(* IEC 61131-3 sources: daoli-st-library/DL_Algo (part 21) *)

(* ---- FB_DL_SelfDischargeScreen.st ---- *)
(*
  FB_DL_SelfDischargeScreen  —  自放电筛分（压降速率 K 值分级 + 温度补偿） / Self-discharge screening by voltage-drop rate grading with temperature compensation
  分类 Category : DL_Algo
  版本 Version  : 1.0.0
  来源 Source   : roadmap-li-p2 — 锂电自放电筛分工站真缺口
  溯源 Origin   : 道莅 clean-room 实现；K 值 = ΔOCV/Δt 与 25 °C 温度补偿为公开自放电筛分算法，未复制任何源码行
  功能 Function : 1) 纯计算子函数 FC_DL_SelfDischargeKCalc 求压降速率
                  K = (fOcvStartV - fOcvEndV) / 静置时长(h)，静置时长按秒换算（除 3600.0 常量）；
                  2) 温度补偿：K25 = K / (1.0 + fTempCoeffPerK × (fTempC - 25.0))，
                  分母绝对值 <= 1.0E-6 返回 -1.0 哨兵（不饱和、不置 0，交主块判故障）；
                  3) 分级：K25 与 fClassAMvPerH / fClassBMvPerH / fClassCMvPerH 比较，
                  越 C 档为 eReject（ELSE 兜底）；
                  4) 报告值向上取整到 0.001 mV/h（先实数上限兜底 → 截断 → 余量进位，
                  正好整除不 +1，禁 TRUNC(x)+1）；
                  5) 本件只有故障码、无信息码（派单硬约束）。
  接口 Interface: 输入首末 OCV/静置时长/温度/温度系数/三档阈值；输出 K/K25/取整值/分级/码
  边界 Boundary : ① 组态闸：tRest <= T#0S、fTempCoeffPerK < 0.0、fClassAMvPerH < 0.0、
                  fClassBMvPerH <= fClassAMvPerH、fClassCMvPerH <= fClassBMvPerH
                  → 0389 锁存；② 首末 OCV 非有限（NaN 自反 + Inf 差值自减）→ 0389 锁存；
                  ③ 温补分母哨兵 -1.0 由主块转 0389 锁存（子函数不置故障）；
                  ④ 取整前实数上限兜底防 LREAL→DINT 溢出；⑤ 仅一个 R_TRIG，段 0 无条件调用；
                  ⑥ 故障相迁出唯一路径 = bReset 上升沿；⑦ 零全局耦合（无 GVL / %I %Q %M）。
  依赖 Depends  : Standard.library（R_TRIG）
  码表 Error codes（Algo 段 0002，故障窗口 0389；本件无信息码）:
    16#0002_0389 故障级：自放电筛分故障总码（组态非法 / OCV 非有限 / 温补分母非法），
                 锁存至 bReset 上升沿；归因见 eCause，不新增码位（派单硬约束单码）
  修订历史 Revision :
    2026-11-19  v1.0.0  R43 首版（批次 3 · 序号 13）
*)

TYPE E_DL_SdsState :
(
    eIdle   := 0,     // 未使能待筛分 / Idle, waiting screening
    eRun    := 10,    // 筛分计算中 / Screening active
    eFault  := 90     // 故障锁存相 / Fault latched phase
);
END_TYPE

TYPE E_DL_SdsClass :
(
    eNone   := 0,     // 未分级 / Not graded
    eClassA := 1,     // A 级（自放电最小） / Class A, lowest self-discharge
    eClassB := 2,     // B 级 / Class B
    eClassC := 3,     // C 级 / Class C
    eReject := 4      // 不合格（越 C 档） / Rejected
);
END_TYPE

TYPE E_DL_SdsCause :
(
    eNone       := 0, // 无故障成因 / No cause
    eCfgIllegal := 1, // 组态非法 / Illegal configuration
    eNonFinite  := 2, // OCV 非有限 / Non-finite OCV
    eCompDiv    := 3  // 温补分母非法 / Invalid compensation denominator
);
END_TYPE

FUNCTION FC_DL_SelfDischargeKCalc : REAL
VAR_INPUT
    fOcvStartV     : REAL;   // 静置前 OCV [V] / OCV before rest
    fOcvEndV       : REAL;   // 静置后 OCV [V] / OCV after rest
    fRestS         : REAL;   // 静置时长 [s]，域 > 0 / Rest duration in seconds
    fTempC         : REAL;   // 电芯温度 [°C] / Cell temperature
    fTempCoeffPerK : REAL;   // 温度系数 [1/K]，域 >= 0 / Temperature coefficient
END_VAR
VAR
    _fKPerH  : REAL;         // 未补偿压降速率 [V/h] / Uncompensated drop rate
    _fDen    : REAL;         // 温补分母 [-] / Compensation denominator
END_VAR
(* 纯计算子函数：K25 = K / (1 + coeff × (T - 25))；分母非法返回 -1.0 哨兵 *)
IF fRestS <= 1.0E-6 THEN                              // 除零前置判（时长正域） / Duration positive check
    FC_DL_SelfDischargeKCalc := -1.0;                 // 哨兵：时长非法 / Sentinel
    RETURN;
END_IF
_fKPerH := (fOcvStartV - fOcvEndV) / (fRestS / 3600.0);   // 压降速率 [V/h]（除常量 3600.0） / Drop rate
_fDen := 1.0 + fTempCoeffPerK * (fTempC - 25.0);          // 温补分母 / Compensation denominator
IF ABS(_fDen) <= 1.0E-6 THEN                          // 分母近零判据 / Near-zero denominator
    FC_DL_SelfDischargeKCalc := -1.0;                 // 哨兵：分母非法 / Sentinel
    RETURN;
END_IF
FC_DL_SelfDischargeKCalc := _fKPerH / _fDen * 1000.0; // 补偿后速率 [mV/h] / Compensated rate
END_FUNCTION

FUNCTION_BLOCK FB_DL_SelfDischargeScreen
VAR_INPUT
    fOcvStartV      : REAL := 0.0;      // 静置前 OCV [V] / OCV before rest
    fOcvEndV        : REAL := 0.0;      // 静置后 OCV [V] / OCV after rest
    tRest           : TIME := T#24H;    // 静置时长 [ms]，域 > 0 / Rest duration
    fTempC          : REAL := 25.0;     // 电芯温度 [°C] / Cell temperature
    fTempCoeffPerK  : REAL := 0.002;    // 温度系数 [1/K]，域 >= 0 / Temperature coefficient
    fClassAMvPerH   : REAL := 0.50;     // A 级上限 [mV/h] / Class A limit
    fClassBMvPerH   : REAL := 1.00;     // B 级上限 [mV/h] / Class B limit
    fClassCMvPerH   : REAL := 2.00;     // C 级上限 [mV/h] / Class C limit
    bEnable         : BOOL := FALSE;    // 筛分使能（电平）[-] / Screening enable
    bReset          : BOOL := FALSE;    // 复位命令，上升沿清故障 [-] / Reset edge
END_VAR
VAR_OUTPUT
    eState          : E_DL_SdsState;    // 状态出口，段 6 单点映射 / State outlet
    eClass          : E_DL_SdsClass;    // 分级出口 / Grading outlet
    eCause          : E_DL_SdsCause;    // 故障成因出口（R190） / Fault cause outlet
    fKMvPerH        : REAL;             // 温补后压降速率 [mV/h] / Compensated drop rate
    fKCeilMvPerH    : REAL;             // 向上取整到 0.001 的速率 [mV/h] / Ceiled rate
    bError          : BOOL;             // 故障锁存标志 [-] / Fault latch flag
    nErrId          : UDINT;            // 故障码，0 = 无故障（本件无信息码） / Fault code only
END_VAR
VAR
    _eState         : E_DL_SdsState := E_DL_SdsState.eIdle;   // 内部相位（CASE 唯一写入目标） / Internal phase
    _eClass         : E_DL_SdsClass := E_DL_SdsClass.eNone;   // 分级槽（每拍重算） / Grading slot
    _eCause         : E_DL_SdsCause := E_DL_SdsCause.eNone;   // 故障成因锁存（锁存量） / Latched cause
    rtReset         : R_TRIG;           // 复位沿实例，每周期无条件调用 / Reset edge
    _fK             : REAL;             // 子函数返回速率 [mV/h]（当拍量） / Sub-function result
    _fScaled        : REAL;             // 取整中间量（×1000 后） / Scaling intermediate
    _iScaled        : DINT;             // 截断后整数（×1000） / Truncated integer
    _bNonFin        : BOOL;             // OCV 非有限当拍量 [-] / Non-finite OCV
    _bCfgBad        : BOOL;             // 组态非法当拍量 [-] / Config illegal
    _bFault         : BOOL;             // 故障锁存位（锁存量） / Latched fault bit
    _uFault         : UDINT;            // 故障码锁存（锁存量） / Latched fault code
END_VAR

(* —— 段 0：沿实例无条件周期刷新 + 当拍量判据 —— *)
_bNonFin := (fOcvStartV <> fOcvStartV) OR (fOcvEndV <> fOcvEndV) OR (fTempC <> fTempC)
         OR ((fOcvStartV - fOcvStartV) <> (fOcvStartV - fOcvStartV))
         OR ((fOcvEndV - fOcvEndV) <> (fOcvEndV - fOcvEndV))
         OR ((fTempC - fTempC) <> (fTempC - fTempC));                        // NaN 自反 + Inf 差值自减 / NaN and Inf
_bCfgBad := (tRest <= T#0S) OR (fTempCoeffPerK < 0.0) OR (fClassAMvPerH < 0.0)
            OR (fClassBMvPerH <= fClassAMvPerH) OR (fClassCMvPerH <= fClassBMvPerH);   // 组态非法当拍量 / Config illegal
rtReset(CLK := bReset);                                                      // 复位沿，每拍必调 / Reset edge

(* —— 段 1：单拍量预清零（锁存量不入清单；分级槽每拍重算） —— *)
eClass := E_DL_SdsClass.eNone;      // 分级出口缺省未分级 / Grading default
fKMvPerH := 0.0;                    // 速率出口缺省 0 / Rate default
fKCeilMvPerH := 0.0;                // 取整出口缺省 0 / Ceil default
nErrId := 16#0000_0000;             // 故障码缺省无故障 / Fault code default

(* —— 段 2：复位沿 + 组态域闸 —— *)
IF rtReset.Q THEN                              // rtReset.Q = 当拍量 / current scan
    _bFault := FALSE;                          // 清故障锁存位（锁存量） / Clear fault latch
    _uFault := 16#0000_0000;                   // 清故障锁存码（锁存量） / Clear fault code
    _eCause := E_DL_SdsCause.eNone;            // 清成因（锁存量） / Clear cause
    IF _eState = E_DL_SdsState.eFault THEN
        _eState := E_DL_SdsState.eIdle;        // 故障相迁出：回未使能 / Fault exit to idle
    END_IF
END_IF
IF _bNonFin THEN                               // 非有限锁存 / Non-finite latch
    _uFault := 16#0002_0389;                   // 故障级：筛分故障总码 / Algo fault code
    _eCause := E_DL_SdsCause.eNonFinite;       // 归因：非有限 / Cause: non-finite
    _bFault := TRUE;                           // 标志与码位配对（R45） / Flag paired with code
END_IF
IF _bCfgBad THEN                               // 组态域闸 / Config gate
    _uFault := 16#0002_0389;
    _eCause := E_DL_SdsCause.eCfgIllegal;      // 归因：组态非法 / Cause: illegal config
    _bFault := TRUE;
END_IF

(* —— 段 3：K 值计算 + 温补哨兵 + 取整 + 分级（仅运行相且无故障） —— *)
IF (NOT _bFault) AND (_eState = E_DL_SdsState.eRun) THEN
    _fK := FC_DL_SelfDischargeKCalc(fOcvStartV := fOcvStartV, fOcvEndV := fOcvEndV,
                                    fRestS := TIME_TO_REAL(tRest) / 1000.0,
                                    fTempC := fTempC, fTempCoeffPerK := fTempCoeffPerK);   // 子函数求解（除零由子函数守卫） / Sub-function call
    IF _fK < 0.0 THEN                                      // 哨兵：时分母或时长非法 / Sentinel from sub-function
        _uFault := 16#0002_0389;
        _eCause := E_DL_SdsCause.eCompDiv;                 // 归因：温补分母非法 / Cause: denominator
        _bFault := TRUE;
    ELSE
        fKMvPerH := _fK;                                   // 速率镜像 / Rate mirror
        _fScaled := _fK * 1000.0;                           // 放大 1000 倍进入整数域 / Scale by thousand
        IF _fScaled >= 2.147483E9 THEN                      // 实数上限兜底（DINT 可表上界） / Real upper guard
            _fScaled := 2.147483E9;
        ELSIF _fScaled <= -2.147483E9 THEN                  // 实数下限兜底 / Real lower guard
            _fScaled := -2.147483E9;
        END_IF
        _iScaled := LREAL_TO_DINT(LREAL(_fScaled));         // 截断取整 / Truncate
        IF LREAL(_iScaled) < LREAL(_fScaled) - 1.0E-9 THEN  // 余量进位（正好整除不进位） / Ceiling by remainder
            _iScaled := _iScaled + 1;
        END_IF
        fKCeilMvPerH := DINT_TO_REAL(_iScaled) * 0.001;     // 还原为 0.001 mV/h 步长 / Restore 0.001 step
        IF fKCeilMvPerH <= fClassAMvPerH THEN
            _eClass := E_DL_SdsClass.eClassA;               // A 级 / Class A
        ELSIF fKCeilMvPerH <= fClassBMvPerH THEN
            _eClass := E_DL_SdsClass.eClassB;               // B 级 / Class B
        ELSIF fKCeilMvPerH <= fClassCMvPerH THEN
            _eClass := E_DL_SdsClass.eClassC;               // C 级 / Class C
        ELSE
            _eClass := E_DL_SdsClass.eReject;               // 不合格（ELSE 兜底） / Rejected fallback
        END_IF
    END_IF
END_IF

(* —— 段 4：故障解除式（R240；全当拍量）：rtReset.Q / NOT _bCfgBad / NOT _bNonFin —— *)
IF rtReset.Q AND (NOT _bCfgBad) AND (NOT _bNonFin) THEN
    _bFault := FALSE;                          // 清故障锁存位（锁存量） / Clear fault latch
    _uFault := 16#0000_0000;                   // 清故障锁存码（锁存量） / Clear fault code
    _eCause := E_DL_SdsCause.eNone;            // 清成因（锁存量） / Clear cause
END_IF

(* —— 段 4A：故障锁存相位迁移闸 —— *)
IF _bFault AND (_eState <> E_DL_SdsState.eFault) THEN
    _eState := E_DL_SdsState.eFault;           // 锁存即入故障相 / Latch enters fault phase
END_IF

(* —— 段 5：相位机（CASE 全覆盖 + ELSE 兜底） —— *)
CASE _eState OF

E_DL_SdsState.eIdle:
    IF bEnable AND (NOT _bFault) THEN          // 使能条件 / Enable gate
        _eState := E_DL_SdsState.eRun;         // 进筛分相 / Enter screening
    END_IF

E_DL_SdsState.eRun:
    IF NOT bEnable THEN                        // 撤使能：回未使能（前置消失） / Disable returns idle
        _eState := E_DL_SdsState.eIdle;
    END_IF

E_DL_SdsState.eFault:
    ;                                          // 故障相：仅段 4 复位沿可迁出 / Only reset exits

ELSE
    _uFault := 16#0002_0389;                   // 故障级：非法相位兜底（归并总码） / Illegal phase fallback
    _eCause := E_DL_SdsCause.eCfgIllegal;      // 归因：相位非法归并组态 / Cause: phase illegal
    _bFault := TRUE;
    _eState := E_DL_SdsState.eFault;           // 强制回故障相 / Force fault phase

END_CASE

(* —— 段 6：出口单点映射（名实同源；锁存码回放） —— *)
IF _bFault THEN
    nErrId := _uFault;                         // 故障锁存码回放 / Replay latched code
    eClass := E_DL_SdsClass.eNone;             // 故障相分级强制未分级 / Grading forced none
    fKCeilMvPerH := 0.0;                       // 故障相取整值强制 0（安全侧） / Ceil forced zero
ELSE
    nErrId := 16#0000_0000;                    // 无故障：本件无信息码 / No fault, no info code
    eClass := _eClass;                         // 分级出口 / Grading outlet
END_IF
bError := _bFault;                             // 故障标志同源 / Flag from latch
eState := _eState;                             // 状态出口 / State outlet
eCause := _eCause;                             // 成因出口 / Cause outlet

END_FUNCTION_BLOCK

(* ---- FB_DL_SensorConsensusSelector.st ---- *)
(*
  FB_DL_SensorConsensusSelector —— 多通道传感器共识选择：中位基准+偏差带剔除+通道不足降级到单通道，ENUM 状态机
  分类：DL_Algo | 复杂度：3 | 轮次：R86
  开源溯源：道莅原创（clean-room 自研，纯 IEC 61131-3 通用算法），无外部代码引用
  许可证：MIT

  职责：对 5 路同类传感器做共识表决——有效通道数 ≥3 时取中位数作基准、剔除超出偏差带的通道后取平均（NORMAL）；
        有效数 =2 取均值、=1 直通（DEGRADED）；有效数 =0 保持上值并置 xLost（LOST）。
  输入契约：arrVal 通道值 [工程单位]；arrValid 通道有效位；fDevBand 偏差带半宽 [工程单位]（> 0）；
            fAbsMax 非有限闸与量程闸的绝对上限 [工程单位]。
  输出契约：fOut 共识值 [工程单位]；nValidOut 参与表决的有效通道数；xValid 本次输出可信；
            xDegraded / xLost 分级标志；eMode 表决模式枚举。
  边界：① 非有限双判（x <> x 判 NaN、ABS(x) > fAbsMax 判 Inf / 越界）逐通道执行；
        ② 除零防护：所有均值前判分母 > 0；③ 排序用插入法（FOR + WHILE 递减），无 FOR..DOWNTO；
        ④ CASE 含 ELSE 兜底把非法模式拦入 LOST；⑤ 零全局耦合、零物理地址、零库件依赖。
*)

(*-----------------------------------------------------------------------------
 * 枚举: E_DL_ConsMode（共识表决模式，归属本文件，全库唯一定义）
 *----------------------------------------------------------------------------*)
TYPE E_DL_ConsMode :
(
    eNormal   := 0,   // 正常共识（≥3 通道且带内 ≥3） [—] / Normal consensus with at least three in band channels
    eDegraded := 1,   // 降级（2 通道均值 / 1 通道直通 / 带内不足 3） [—] / Degraded consensus
    eLost     := 2    // 失效（零有效通道，保持上值） [—] / Lost, holds the previous value
);
END_TYPE

FUNCTION_BLOCK FB_DL_SensorConsensusSelector
VAR_INPUT
    xEnable  : BOOL  := TRUE;                             // 使能，FALSE 时按失效模式处理 [—] / Enable, false is treated as lost
    arrVal   : ARRAY[0..4] OF REAL;                       // 五路通道采样值 [工程单位] / Five channel samples
    arrValid : ARRAY[0..4] OF BOOL;                       // 五路通道有效位 [—] / Five channel validity flags
    fDevBand : REAL  := 1.0;                              // 偏差带半宽，必须 > 0 [工程单位] / Deviation band half width
    fAbsMax  : REAL  := 1.0E30;                           // 数值绝对上限（非有限 / 越界闸） [工程单位] / The absolute magnitude gate
END_VAR
VAR_OUTPUT
    fOut       : REAL;                                    // 共识输出值 [工程单位] / The consensus output value
    nValidOut  : INT;                                     // 参与表决的有效通道数 [个] / The number of channels taking part
    xValid     : BOOL;                                    // 本次输出可信 [—] / The output is trustworthy
    xDegraded  : BOOL;                                    // 降级标志 [—] / The degraded flag
    xLost      : BOOL;                                    // 失效标志 [—] / The lost flag
    eMode      : E_DL_ConsMode;                           // 表决模式枚举 [—] / The consensus mode enumeration
END_VAR
VAR
    afSort    : ARRAY[0..4] OF REAL;                      // 有效值排序缓冲（升序） [工程单位] / The ascending sort buffer
    nCnt      : INT;                                      // 有效通道数 [个] / The valid channel count
    nIn       : INT;                                      // 偏差带内通道数 [个] / The in band channel count
    k         : INT;                                      // 外层遍历索引 [下标] / The outer loop index
    j         : INT;                                      // 插入排序内层索引 [下标] / The insertion sort index
    fTmp      : REAL;                                     // 插入排序暂存量 [工程单位] / The insertion sort temporary
    fMed      : REAL;                                     // 中位数基准 [工程单位] / The median reference
    fSum      : REAL;                                     // 带内累加和 [工程单位] / The in band accumulation
    fMean     : REAL;                                     // 带内均值 [工程单位] / The in band mean
    fCand     : REAL;                                     // 候选输出值 [工程单位] / The candidate output value
    fDiff     : REAL;                                     // 单通道与中位数的偏差 [工程单位] / The deviation from the median
    fLastOut  : REAL;                                     // 上拍共识输出保持量 [工程单位] / The held previous output
    xHasLast  : BOOL;                                     // 是否已有可用上拍值 [—] / Whether a previous value exists
    eCand     : E_DL_ConsMode;                            // 候选表决模式 [—] / The candidate mode
END_VAR
VAR CONSTANT
    DL_CM_ZERO : INT := 0;                                // 整型零常量 [个] / The integer zero constant
    DL_CM_ONE  : INT := 1;                                // 整型一常量 [个] / The integer one constant
    DL_CM_NCH  : INT := 5;                                // 通道总数 [个] / The total channel count
    DL_CM_MINC : INT := 3;                                // 正常共识所需最少通道数 [个] / The minimum channels for normal consensus
    DL_CM_R0   : REAL := 0.0;                             // 浮点零常量 [工程单位] / The floating point zero constant
    DL_CM_EPS  : REAL := 1.0E-6;                          // 浮点比较容差 [工程单位] / The floating point comparison tolerance
END_VAR

// 段 1｜输出预置（单点预置，CASE 之后不再无条件清零）
xValid := FALSE;                                          // 可信位预置假 / preset the valid flag false
xDegraded := FALSE;                                       // 降级位预置假 / preset the degraded flag false
xLost := FALSE;                                           // 失效位预置假 / preset the lost flag false
nValidOut := DL_CM_ZERO;                                  // 有效通道数预置零 [个] / preset the valid count zero
nCnt := DL_CM_ZERO;                                       // 排序缓冲计数预置零 [个] / preset the buffer count zero
fMed := DL_CM_R0;                                         // 中位数预置零 [工程单位] / preset the median zero
fCand := fLastOut;                                        // 候选值默认继承上拍值 [工程单位] / default the candidate to the held value

// 段 2｜逐通道有效性 + 非有限闸，有效值收集进排序缓冲
FOR k := DL_CM_ZERO TO DL_CM_NCH - 1 DO                   // 五通道遍历（上界 4 已由常量钉死） / traverse all channels
    IF arrValid[k] THEN                                   // 通道有效位为真 / the channel is flagged valid
        IF (arrVal[k] <> arrVal[k]) THEN                  // 自反判 NaN / the self comparison catches NaN
            fTmp := DL_CM_R0;                             // 置暂存零（本通道将被剔除） / stage zero, channel dropped
        ELSIF ABS(arrVal[k]) > fAbsMax THEN               // 越绝对上限判 Inf / 越界 / beyond the magnitude gate
            fTmp := DL_CM_R0;                             // 置暂存零（本通道将被剔除） / stage zero, channel dropped
        ELSE
            afSort[nCnt] := arrVal[k];                    // 有效值入缓冲 [工程单位] / store the valid value
            nCnt := nCnt + DL_CM_ONE;                     // 有效计数自增 [个] / increment the valid count
        END_IF
    END_IF
END_FOR
nValidOut := nCnt;                                        // 有效通道数出口 [个] / publish the valid count

// 段 3｜插入排序升序（WHILE 显式递减，禁 FOR..DOWNTO）
FOR k := DL_CM_ONE TO nCnt - DL_CM_ONE DO                 // 从第二个元素起逐个插入 / insert every element from the second
    IF k >= DL_CM_ONE THEN                                // k 合法且缓冲至少有 k+1 个元素 / k is legal with enough elements
        fTmp := afSort[k];                                // 取出待插入元素 [工程单位] / take the element to insert
        j := k - DL_CM_ONE;                               // 内层索引从 k-1 起 / the inner index starts at k minus one
        WHILE (j >= DL_CM_ZERO) AND (afSort[j] > fTmp) DO // 显式递减并判下界 / explicit decrement with a bound check
            afSort[j + DL_CM_ONE] := afSort[j];           // 逆序元素右移一格 / shift the larger element right
            j := j - DL_CM_ONE;                           // 内层索引递减 [下标] / decrement the inner index
        END_WHILE
        afSort[j + DL_CM_ONE] := fTmp;                    // 待插入元素落位 [工程单位] / land the element
    END_IF
END_FOR

// 段 4｜按有效通道数分档：中位数基准 + 偏差带剔除 + 候选模式判定
IF (NOT xEnable) OR (nCnt = DL_CM_ZERO) THEN              // 未使能或零有效通道 / disabled or no valid channel
    eCand := E_DL_ConsMode.eLost;                         // 候选模式判失效 / the candidate mode is lost
ELSIF nCnt = DL_CM_ONE THEN                               // 单通道直通 / a single channel passes through
    fCand := afSort[0];                                   // 直通该通道值 [工程单位] / pass the single value
    eCand := E_DL_ConsMode.eDegraded;                     // 候选模式判降级 / the candidate mode is degraded
ELSIF nCnt = DL_CM_ONE + DL_CM_ONE THEN                   // 双通道取均值 / two channels take the mean
    fCand := (afSort[0] + afSort[1]) / 2.0;               // 双通道均值 [工程单位] / the mean of the two channels
    eCand := E_DL_ConsMode.eDegraded;                     // 候选模式判降级 / the candidate mode is degraded
ELSE                                                      // 三通道及以上做中位基准表决 / three or more channels vote
    IF (nCnt MOD 2) = DL_CM_ONE THEN                      // 奇数个取正中位 / odd count takes the middle element
        fMed := afSort[nCnt / 2];                         // 中位数基准 [工程单位] / the median reference
    ELSE
        fMed := (afSort[nCnt / 2 - DL_CM_ONE] + afSort[nCnt / 2]) / 2.0; // 偶数个取中间两值均值 [工程单位]
    END_IF
    nIn := DL_CM_ZERO;                                    // 带内计数清零 [个] / clear the in band count
    fSum := DL_CM_R0;                                     // 带内和清零 [工程单位] / clear the in band sum
    FOR k := DL_CM_ZERO TO nCnt - DL_CM_ONE DO             // 遍历有效通道做偏差带剔除 / filter by the deviation band
        fDiff := afSort[k] - fMed;                        // 与中位数的偏差 [工程单位] / the deviation from the median
        IF ABS(fDiff) <= fDevBand THEN                    // 带内（含边界，容差口径） / inside the band
            fSum := fSum + afSort[k];                     // 累加带内值 [工程单位] / accumulate the in band value
            nIn := nIn + DL_CM_ONE;                       // 带内计数自增 [个] / increment the in band count
        END_IF
    END_FOR
    IF nIn >= DL_CM_MINC THEN                             // 带内至少 3 通道 / at least three channels stay in band
        fMean := fSum / INT_TO_REAL(nIn);                 // 带内均值（分母 ≥3 已证非零） [工程单位] / the in band mean
        fCand := fMean;                                   // 候选输出取带内均值 [工程单位] / the candidate is the mean
        eCand := E_DL_ConsMode.eNormal;                    // 候选模式判正常 / the candidate mode is normal
    ELSIF nIn = DL_CM_ONE + DL_CM_ONE THEN                // 带内仅剩 2 通道 / only two channels stay in band
        fMean := fSum / 2.0;                              // 两通道均值 [工程单位] / the mean of the two channels
        fCand := fMean;                                   // 候选输出取该均值 [工程单位] / the candidate is that mean
        eCand := E_DL_ConsMode.eDegraded;                 // 候选模式判降级 / the candidate mode is degraded
    ELSE                                                  // 带内不足 2 通道，退回中位基准 / too few in band, fall back to the median
        fCand := fMed;                                    // 候选输出取中位数 [工程单位] / the candidate is the median
        eCand := E_DL_ConsMode.eDegraded;                 // 候选模式判降级 / the candidate mode is degraded
    END_IF
END_IF

// 段 5｜模式出口分派（ENUM + CASE，ELSE 拦截非法模式）
CASE eCand OF
    E_DL_ConsMode.eNormal:
        fOut := fCand;                                    // 正常模式直接输出候选值 [工程单位] / publish the candidate
        xValid := TRUE;                                   // 置可信位 [—] / raise the valid flag
        xDegraded := FALSE;                               // 清降级位 [—] / clear the degraded flag
        xLost := FALSE;                                   // 清失效位 [—] / clear the lost flag
        fLastOut := fOut;                                 // 刷新保持量 [工程单位] / refresh the held value
        xHasLast := TRUE;                                 // 保持量可用 [—] / the held value is now available
    E_DL_ConsMode.eDegraded:
        fOut := fCand;                                    // 降级模式输出候选值 [工程单位] / publish the candidate
        xValid := TRUE;                                   // 降级输出仍可信 [—] / a degraded output is still valid
        xDegraded := TRUE;                                // 置降级位 [—] / raise the degraded flag
        xLost := FALSE;                                   // 清失效位 [—] / clear the lost flag
        fLastOut := fOut;                                 // 刷新保持量 [工程单位] / refresh the held value
        xHasLast := TRUE;                                 // 保持量可用 [—] / the held value is now available
    E_DL_ConsMode.eLost:
        IF xHasLast THEN                                  // 已有上拍值 / a previous value exists
            fOut := fLastOut;                             // 保持上拍值 [工程单位] / hold the previous value
        ELSE
            fOut := DL_CM_R0;                             // 无上拍值输出零哨兵 [工程单位] / zero sentinel without history
        END_IF
        xValid := FALSE;                                  // 失效输出不可信 [—] / the lost output is not valid
        xDegraded := TRUE;                                // 失效同时视为降级 [—] / lost is also degraded
        xLost := TRUE;                                    // 置失效位 [—] / raise the lost flag
ELSE
    fOut := DL_CM_R0;                                     // 非法模式输出零哨兵 [工程单位] / illegal mode outputs the zero sentinel
    xValid := FALSE;                                      // 非法模式不可信 [—] / an illegal mode is not valid
    xDegraded := TRUE;                                    // 非法模式视为降级 [—] / an illegal mode is degraded
    xLost := TRUE;                                        // 非法模式视为失效 [—] / an illegal mode is lost
    eCand := E_DL_ConsMode.eLost;                          // 非法模式回写为失效 [—] / normalise the illegal mode to lost
END_CASE
eMode := eCand;                                           // 模式枚举单点出口 / the single point mode outlet
END_FUNCTION_BLOCK

(* ---- FB_DL_SensorDriftBaseline.st ---- *)
(*
  Name        : FB_DL_SensorDriftBaseline
  Category    : DL_Algo
  Version     : 1.0.1
  Purpose     : 传感器慢漂移基线跟踪：长窗指数（EMA）基线随测量缓慢跟随，测量对基线的快偏差超限经确认延时即报警（区分真实工况阶跃与传感器漂移）；/ Sensor slow-drift baseline tracking: a long-window EMA baseline follows the measurement, and a fast deviation beyond limit confirmed over a delay raises an alarm
  溯源        : 借 t2-1-measurement 的分类/参数域组织，clean-room 实现
  Changelog   : v1.0.1 R54 非有限输入穿透修复：迁入拍/基线更新/残差出口前置有限性闸，非有限拍冻结基线并置 bSensorBad，出口保持上拍值
  Boundary    : ① 组态闸：基线因子域 (0..1] / 快偏差限 > 0 / 确认延时 > 0 → 锁存故障（因子 0/1 端点使基线冻结或退化为直通）；
                ② 非有限测量该拍不更新基线（基线保持上拍值，防污染慢积分器），判据整拍跳过；
                ③ 基线快照在迁入 eMon 拍取（fValue 首值），避免从 0 慢爬造成的假偏差；
                ④ 确认延时 TON 串 eMon 相位闸（族③），段 0 无 IF 包裹；
                ⑤ bDriftFast 锁存至复位沿；fBaseline/fDeviation 出口在 eIdle/eFault 有确定值；
                ⑥ 本件为诊断层，不修正测量值、不重标定（属主边界）。
*)
TYPE E_DL_SdbState :
(
    eIdle  := 0,                             (* 未使能 / Disabled *)
    eMon   := 10,                            (* 基线跟踪运行 / Tracking *)
    eFault := 90                             (* 故障锁存相 / Fault latched *)
);
END_TYPE

TYPE E_DL_SdbCause :
(
    eNone       := 0,                        (* 无故障成因 / No cause *)
    eCfgIllegal := 1,                        (* 组态非法：因子/偏差限/延时越域 / Illegal config *)
    eDriftFast  := 2,                        (* 快偏差确认（基线失跟或真实阶跃，上层判别） / Fast deviation confirmed *)
    ePhaseBad   := 3                         (* 非法相位兜底 / Illegal phase fallback *)
);
END_TYPE

FUNCTION_BLOCK FB_DL_SensorDriftBaseline
VAR_INPUT
    fValue    : REAL := 0.0;                 (* 传感器测量值（任意工程量）[-] / Sensor measurement *)
    fAlpha    : REAL := 0.005;               (* 基线 EMA 因子（每拍跟随比例），域 (0..1] [-] / Baseline EMA factor *)
    fFastLim  : REAL := 5.0;                 (* 快偏差报警限，域 > 0 [工程单位] / Fast-deviation limit, > 0 *)
    tConfirm  : TIME := T#30S;               (* 快偏差确认延时，域 > T#0S [ms] / Deviation confirm delay, > 0 *)
    bEnable   : BOOL := TRUE;                (* 跟踪使能 [-] / Enable *)
    bReset    : BOOL := FALSE;               (* 复位命令，上升沿清报警与基线 [-] / Reset command *)
END_VAR
VAR_OUTPUT
    fBaseline : REAL;                        (* 慢漂移基线（EMA 跟踪值）[工程单位] / Slow-drift baseline *)
    fDeviation: REAL;                        (* 测量对基线快偏差（实时派生）[工程单位] / Fast deviation versus baseline *)
    bDriftFast: BOOL;                        (* 快偏差报警锁存（复位沿清）[-] / Fast-deviation alarm latched *)
    bSensorBad: BOOL;                        (* 测量非有限传感器失效锁存（复位沿清，v1.0.1）[-] / Sensor bad latched *)
    eState    : E_DL_SdbState;               (* 状态出口 / State outlet *)
    eCause    : E_DL_SdbCause;               (* 故障成因出口（R190 归因唯一） / Fault cause outlet *)
    bError    : BOOL;                        (* 故障锁存标志 [-] / Fault latch flag *)
END_VAR
VAR
    _eState  : E_DL_SdbState := E_DL_SdbState.eIdle;     (* 内部相位（CASE 唯一写入目标） / Internal phase *)
    _eCause  : E_DL_SdbCause := E_DL_SdbCause.eNone;     (* 故障成因锁存量 / Latched cause *)
    rtReset  : R_TRIG;                       (* 复位沿实例，段 0 无条件调用 / Reset edge instance *)
    tonConf  : TON;                          (* 快偏差确认延时计时器（IN 由偏差判据派生 + 相位闸） / Deviation confirm timer *)
    _bFault  : BOOL;                         (* 故障锁存位 / Latched fault bit *)
    _bCfgBad : BOOL;                         (* 组态非法当拍量 / Illegal config this scan *)
    _bFin    : BOOL;                         (* 测量值有限性当拍量 / Measurement finiteness *)
    _bBase   : BOOL;                         (* 基线已建立标志 / Baseline established flag *)
    _fBaseI  : REAL;                         (* 基线内部量（EMA 状态）[工程单位] / Baseline internal EMA state *)
    _fDevI   : REAL;                         (* 快偏差中间量 [工程单位] / Deviation intermediate *)
    _fDevLast: REAL;                         (* 上拍有效偏差快照（非有限拍出口冻结用，v1.0.1）[工程单位] / Last valid deviation snapshot *)
    _bDevRaw : BOOL;                         (* 快偏差原始判据当拍量 / Raw deviation verdict *)
END_VAR
VAR CONSTANT
    DL_SDB_EPS  : REAL := 1.0E-6;            (* 判零容差 [-] / Epsilon *)
    DL_SDB_ONE  : REAL := 1.0;               (* 因子上界常量 [-] / Factor upper bound *)
END_VAR

(* —— 段 0：当拍判据派生 + 实例无条件刷新（R228A；R_TRIG/TON 全在段 0，无 IF 包裹） —— *)
_bCfgBad := (fAlpha <= DL_SDB_EPS) OR (fAlpha > DL_SDB_ONE)                    (* 基线因子域闸 (0..1]（端点退化解拦截） / Factor domain gate *)
            OR (fFastLim <= DL_SDB_EPS)                                        (* 快偏差限正域闸 / Deviation limit gate *)
            OR NOT (tConfirm > T#0S);                                          (* 确认延时正域闸 / Confirm delay gate *)
rtReset(CLK := bReset);                                                        (* 复位沿每拍必调 / Reset edge every scan *)
_bFin := (fValue = fValue) AND ((fValue - fValue) = (fValue - fValue));        (* 测量值 NaN 自反 + Inf 差判闸 / Measurement NaN and Inf gate *)
_fDevI := 0.0;                                                                 (* 偏差中间量预置（基线无效期为 0，不误触发计时） / Deviation preset zero *)
IF _bFin AND _bBase THEN
    _fDevI := fValue - _fBaseI;                                                (* 快偏差 = 测量 - 基线（基线已建立才派生）[工程单位] / Deviation versus baseline *)
END_IF
_bDevRaw := _bFin AND _bBase AND (ABS(_fDevI) > fFastLim);                     (* 原始判据：有限 + 基线在 + 超限（直比阈值，非浮点等值） / Raw deviation verdict *)
tonConf(IN := (_eState = E_DL_SdbState.eMon) AND _bDevRaw, PT := tConfirm);    (* 确认延时：判据持续才计时，串 eMon 相位闸 / Confirm timer with phase gate *)

(* —— 段 1：单拍量预清零（R107；bDriftFast 为锁存出口不预清，复位沿清，族② 口径） —— *)
fBaseline := 0.0;                                                              (* 基线出口预清（派生拍覆盖） / Baseline outlet preset *)
fDeviation := 0.0;                                                             (* 偏差出口预清 / Deviation outlet preset *)

(* —— 段 2：复位沿处理（作用域：清故障 + 清报警 + 清基线 + 迁 eIdle，R283 逐项声明） —— *)
IF rtReset.Q THEN
    _bFault := FALSE;                                                          (* 清故障锁存 / Clear fault *)
    _eCause := E_DL_SdbCause.eNone;                                            (* 清成因 / Clear cause *)
    bDriftFast := FALSE;                                                       (* 清快偏差报警锁存 / Clear alarm latch *)
    _bBase := FALSE;                                                           (* 清基线已建立位（重使能重新取快照） / Clear baseline flag *)
    _fBaseI := 0.0;                                                            (* 清基线内部量 / Clear baseline internal *)
    _fDevLast := 0.0;                                                          (* 清有效偏差快照（v1.0.1） / Clear deviation snapshot *)
    bSensorBad := FALSE;                                                       (* 清传感器失效锁存（v1.0.1） / Clear sensor bad latch *)
    fBaseline := 0.0;                                                          (* 清基线出口 / Clear baseline outlet *)
    fDeviation := 0.0;                                                         (* 清偏差出口 / Clear deviation outlet *)
    _eState := E_DL_SdbState.eIdle;                                            (* 迁未使能相 / Back to idle *)
END_IF

(* —— 段 3：组态故障锁存（锁存至复位沿，R189） —— *)
IF _bCfgBad AND NOT _bFault THEN
    _bFault := TRUE;                                                           (* 锁存故障位 / Latch fault *)
    _eCause := E_DL_SdbCause.eCfgIllegal;                                      (* 成因：组态非法 / Cause: illegal config *)
    _eState := E_DL_SdbState.eFault;                                           (* 同步迁故障相 / Migrate to fault *)
END_IF

(* —— 段 4：CASE 主状态机（ELSE 兜底迁 eFault，红线 6） —— *)
CASE _eState OF
    E_DL_SdbState.eIdle:                                                       (* 未使能：出口确定值 / Disabled *)
        fBaseline := 0.0;                                                      (* 失能清基线出口 / Clear baseline outlet *)
        fDeviation := 0.0;                                                     (* 失能清偏差出口 / Clear deviation outlet *)
        bDriftFast := FALSE;                                                   (* 失能清报警出口 / Clear alarm outlet *)
        _bBase := FALSE;                                                       (* 失能清基线位（重使能重新对齐） / Clear baseline flag *)
        bSensorBad := FALSE;                                                   (* 失能清传感器失效出口（确定值） / Clear sensor bad *)
        IF bEnable AND NOT _bFault AND _bFin THEN                              (* 迁入闸加有限性闸：迁入拍为非有限不建基线不迁入（v1.0.1 修复） / Entry gate with finiteness *)
            _fBaseI := fValue;                                                 (* 迁入拍取基线首快照（相位闸配套，边界③） / Baseline snapshot at entry *)
            _bBase := TRUE;                                                    (* 基线已建立 / Baseline established *)
            _eState := E_DL_SdbState.eMon;                                     (* 使能进入跟踪 / Enter tracking *)
        END_IF
    E_DL_SdbState.eMon:                                                        (* 跟踪相：EMA 基线 + 快偏差判 / Tracking *)
        IF NOT bEnable THEN
            _eState := E_DL_SdbState.eIdle;                                    (* 失能回未使能 / Back to idle *)
        ELSE
            fBaseline := _fBaseI;                                              (* 基线出口（状态镜像，R191；非有限拍 _fBaseI 冻结即保持上拍） / Baseline outlet *)
            IF _bFin THEN
                fDeviation := _fDevI;                                          (* 偏差出口（有限拍派生） / Deviation outlet *)
                _fDevLast := _fDevI;                                           (* 有效偏差快照推进（v1.0.1） / Advance deviation snapshot *)
                _fBaseI := _fBaseI + fAlpha * (fValue - _fBaseI);              (* EMA 基线慢跟随（因子域闸保证 (0..1]） / EMA baseline update *)
            ELSE
                fDeviation := _fDevLast;                                       (* 非有限拍：偏差出口保持上拍值（v1.0.1 修复） / Hold last deviation *)
                bSensorBad := TRUE;                                            (* 非有限拍置传感器失效锁存（复位沿清，v1.0.1） / Sensor bad latch *)
            END_IF
            IF tonConf.Q THEN                                                  (* 快偏差持续满确认延时：报警 / Deviation confirmed *)
                bDriftFast := TRUE;                                            (* 报警锁存（复位沿清） / Latch alarm *)
                _bFault := TRUE;                                               (* 同步故障锁存（R45 配对） / Latch fault *)
                _eCause := E_DL_SdbCause.eDriftFast;                           (* 成因：快偏差 / Cause: fast deviation *)
            END_IF
        END_IF
    E_DL_SdbState.eFault:                                                      (* 故障相：冻结保持末值，仅复位沿出 / Fault *)
        ;                                                                      (* 锁存回放（R28） / Replay from latch *)
    ELSE                                                                       (* 非法相位兜底迁安全态 / Illegal phase fallback *)
        _eState := E_DL_SdbState.eFault;                                       (* 迁故障相 / To fault *)
        _bFault := TRUE;                                                       (* 同步锁存 / Latch *)
        _eCause := E_DL_SdbCause.ePhaseBad;                                    (* 成因：非法相位 / Cause: illegal phase *)
END_CASE

(* —— 段 5：出口映射（bError/eState 同源，R191） —— *)
bError := _bFault;                                                             (* 故障标志镜像 / Fault flag mirror *)
eState := _eState;                                                             (* 状态出口 / State outlet *)
eCause := _eCause;                                                             (* 成因出口 / Cause outlet *)
END_FUNCTION_BLOCK

(* ---- FB_DL_SensorFusion2.st ---- *)
(*==============================================================================
 * 组件名称 (Component)  : FB_DL_SensorFusion2
 * 所属子库 (Sublibrary) : DL_Algo
 * 当前版本 (Version)    : 1.0.1
 * 兼容性   (Platform)   : CODESYS 3.5+ / TwinCAT 3 / 汇川 InoProShop / 施耐德 Machine Expert
 *                         仅依赖 Standard.library（ABS），零厂商私有库
 * 功能描述 (Function)   : 双传感器方差加权融合：对同一物理量的两路测量（如 RTD+红外温漂
 *                         互补型双测）按在线递推噪声方差倒数动态配权：
 *                           _fVarX := (1-fTauVar)×_fVarX + fTauVar×(fMeasX-_fMean)²
 *                           fWeightA = (1/_fVarA) / ((1/_fVarA)+(1/_fVarB))
 *                           fFused   = fWeightA×fMeasA + (1-fWeightA)×fMeasB
 *                         一致性判据 bAgree = |fMeasA-fMeasB| <= fDevMax；单源失效全权重
 *                         交给健康源（降级不拒算）；双源失效冻结上次 fFused 且 bValid=FALSE。
 * 接口     (Interface)  : 输入 fMeasA/fMeasB 双路测量、bFreshA/bFreshB 数据新鲜度、
 *                         fTauVar 方差递推平滑系数（域 0~1 无量纲）、fDevMax 一致性偏差闸
 *                         （工程单位）、bReset 复位；输出 fFused 融合值、fWeightA 权重
 *                         （0~1）、bAgree 一致性、bValid 有效标志、bError 故障标志。
 * 边界     (Boundary)   : ① **属主边界（写死）：本件只做双源静态融合，不判传感器硬故障、
 *                         不切换通道、不接管信号健康诊断**；通道硬失效裁决归
 *                         `FB_DL_RedundantSwitch`（二选一切换），本件是"都信、按噪声配权"。
 *                         ② 方差下限钳 fVarMin（VAR CONSTANT）防除零：权重分母两项各含
 *                         1/_fVarX，钳底后分母恒正，无需额外除零判。
 *                         ③ 非有限值当拍剔除（R245）：该源当拍视同不新鲜；双源当拍均剔除
 *                         → 冻结 fFused、bValid=FALSE。
 *                         ④ 权重输出钳 [0,1]；fTauVar 组态域闸（<0 或 >1）与 fDevMax<0
 *                         → 锁存 bError，冻结输出，解除沿 = bReset 上升沿。
 *                         ⑤ 方差递推仅在双源同拍有效时进行（单源降级只直通，不污染方差）。
 *                         ⑥ 零全局耦合（无 GVL / 无 VAR_EXTERNAL / 无物理地址）。
 * 分工声明 (Scope)      : 与 `FB_DL_KalmanFilter1D` 分工：单流递推滤波 ≠ 双源加权融合；
 *                         与 `FB_DL_RedundantSwitch` 分工：二选一切换 ≠ 加权融合（见①）。
 * 来源标签 (Source Tag) : 自研线（公开加权融合公式 clean-room，逆方差权重为公开统计定义）
 * 码表     (Codes)      : 本件不占用任何全局数字码位。出口为 LREAL 组 + BOOL 组；
 *                         数字码位待主控收口阶段统一派号。
 * 红线自检 (Redline)    : R1 ✓ 零 GVL/VAR_EXTERNAL ｜ R2 ✓ 零 %I/%Q/%M ｜ R3 ✓ 纯 IEC 61131-3
 *                         R4 ✓ 方差下限防除零 + 非有限剔除 + 权重钳位 ｜ R5 ✓ 声明逐行同行双语注释
 *                         R6 N/A（无 ENUM 状态机） ｜ R7 ✓ 一 R_TRIG 段 0 无条件刷新
 * 修订历史 (Revision)   : 2026-11-20  v1.0.1  R50 返修 R3：fTauVar=0 端点防护
 *                         （下限钳位）——fTauVar=0 时方差递推步长为零，方差
 *                         永冻结于初值 1.0、权重恒 0.5（自适应失效），现引入
 *                         DL_SF2_TAUMIN(1E-6) 下限钳位使递推保持最低活跃度；
 *                         行为变更同步更新验收向量（fTauVar=0 按 1E-6 生效）。
 *                         2026-11-20  v1.0.0  R48 首版（批次 2 · 序号 6）
 *                         验收向量：等方差双源 → 权重 0.5；A 方差骤增 → 权重移向 B；
 *                         A 不新鲜 → 权重 1.0 全信 B；双源失效 → 冻结 + bValid=FALSE。
 *==============================================================================*)

FUNCTION_BLOCK FB_DL_SensorFusion2
VAR_INPUT
    fMeasA  : LREAL := 0.0;    // A 源测量值 [工程单位] / Source A measurement
    fMeasB  : LREAL := 0.0;    // B 源测量值（与 A 同物理量） [工程单位] / Source B measurement, same quantity as A
    bFreshA : BOOL := TRUE;    // A 源数据新鲜度 [-] / Source A freshness
    bFreshB : BOOL := TRUE;    // B 源数据新鲜度 [-] / Source B freshness
    fTauVar : LREAL := 0.1;    // 方差递推平滑系数，域 [0,1] [无量纲] / Variance recursion smoothing factor
    fDevMax : LREAL := 1.0;    // 一致性偏差闸（|A-B| 超此值 bAgree=FALSE） [工程单位] / Agreement deviation gate
    bReset  : BOOL := FALSE;   // 复位，上升沿清组态故障锁存 [-] / Reset, rising edge clears config fault
END_VAR
VAR_OUTPUT
    fFused   : LREAL;          // 融合输出值 [工程单位] / Fused output value
    fWeightA : LREAL;          // A 源权重，域 [0,1] [-] / Source A weight in [0,1]
    bAgree   : BOOL;           // 双源一致性（单源降级恒 TRUE） [-] / Two-source agreement
    bValid   : BOOL;           // 融合有效标志（双源失效/组态故障为 FALSE） [-] / Fusion validity flag
    bError   : BOOL;           // 组态故障标志（锁存） [-] / Configuration fault flag, latched
END_VAR
VAR
    _fVarA    : LREAL := 1.0;  // A 源在线递推噪声方差（初值 1.0，量纲平方） / Source A recursive noise variance
    _fVarB    : LREAL := 1.0;  // B 源在线递推噪声方差（初值 1.0） / Source B recursive noise variance
    _fMean    : LREAL := 0.0;  // 上拍融合均值（方差递推参考点，冻结源） / Previous fused mean, recursion reference
    _fW       : LREAL := 0.5;  // 当拍权重中间量（冻结源，与出口同源） / Weight intermediate, frozen source
    _fTauUse  : LREAL;         // 生效递推系数（下限钳位后，v1.0.1 端点防护） [-] / Effective smoothing factor after floor clamp
    _fFused   : LREAL := 0.0;  // 融合值锁存镜像（冻结语义源） / Fused value latch mirror
    _bValid   : BOOL;          // 有效标志内部量 / Validity internal
    _bErrLatch: BOOL;          // 组态故障锁存位（解除沿 = bReset 上升沿） / Latched config fault, cleared by reset edge
    rtReset   : R_TRIG;        // 复位沿实例，段 0 无条件调用 / Reset edge instance
    _bUseA    : BOOL;          // A 源当拍可用（新鲜 ∧ 有限） / Source A usable this scan
    _bUseB    : BOOL;          // B 源当拍可用 / Source B usable this scan
    _fInvA    : LREAL;         // A 源逆方差中间量 / Inverse variance of A
    _fInvB    : LREAL;         // B 源逆方差中间量 / Inverse variance of B
    _fDevA    : LREAL;         // A 源对均值偏差 [工程单位] / Deviation of A from mean
    _fDevB    : LREAL;         // B 源对均值偏差 [工程单位] / Deviation of B from mean
END_VAR
VAR CONSTANT
    DL_SF2_VARMIN : LREAL := 1.0E-12;   // 方差下限钳（防除零） [工程单位²] / Variance floor against zero division
    DL_SF2_TAUMIN : LREAL := 1.0E-6;    // 递推系数下限钳（fTauVar=0 端点防护，v1.0.1） [-] / Smoothing factor floor, endpoint guard
    DL_SF2_EPS    : LREAL := 0.0;       // 非有限差值判零基准 [-] / Non-finite difference zero base
    DL_SF2_ONE    : LREAL := 1.0;       // 单位常量（权重钳上限） [-] / Unit constant, weight ceiling
END_VAR

(* —— 段 0：非有限判 + 组态闸 + 沿刷新 —— *)
_bUseA := bFreshA AND (fMeasA = fMeasA) AND ((fMeasA - fMeasA) = DL_SF2_EPS);   // A 源新鲜 ∧ 有限（NaN 自不等 / Inf 差非零，R245） / A fresh and finite
_bUseB := bFreshB AND (fMeasB = fMeasB) AND ((fMeasB - fMeasB) = DL_SF2_EPS);   // B 源新鲜 ∧ 有限 / B fresh and finite
IF (fTauVar < 0.0) OR (fTauVar > DL_SF2_ONE) OR (fDevMax < 0.0) THEN
    _bErrLatch := TRUE;                                    // 组态域闸：锁存（R188 解除沿 = bReset 上升沿） / Config domain gate: latch
END_IF
_fTauUse := fTauVar;                                       // 生效递推系数工作副本 / Effective factor working copy
IF _fTauUse < DL_SF2_TAUMIN THEN
    _fTauUse := DL_SF2_TAUMIN;                             // fTauVar=0 端点钳位：递推保持最低活跃度（v1.0.1） / Endpoint floor clamp
END_IF
rtReset(CLK := bReset);                                    // 复位沿，每拍必调 / Reset edge, every scan

(* —— 段 1：复位沿 —— *)
IF rtReset.Q THEN
    _bErrLatch := FALSE;                                   // 清组态故障锁存 / Clear config fault latch
END_IF

(* —— 段 2：融合主算（组态故障期冻结不重算） —— *)
bValid := FALSE;                                           // 有效标志当拍预清 / Validity preset
IF NOT _bErrLatch THEN
    IF _bUseA AND _bUseB THEN
        _fDevA := fMeasA - _fMean;                         // A 源对上拍均值偏差 / Deviation of A
        _fDevB := fMeasB - _fMean;                         // B 源对上拍均值偏差 / Deviation of B
        _fVarA := (DL_SF2_ONE - _fTauUse) * _fVarA + _fTauUse * _fDevA * _fDevA;   // A 方差递推（生效系数下限钳位后） / A variance recursion
        _fVarB := (DL_SF2_ONE - _fTauUse) * _fVarB + _fTauUse * _fDevB * _fDevB;   // B 方差递推 / B variance recursion
        IF _fVarA < DL_SF2_VARMIN THEN
            _fVarA := DL_SF2_VARMIN;                       // 方差下限钳（防除零） / Variance floor
        END_IF
        IF _fVarB < DL_SF2_VARMIN THEN
            _fVarB := DL_SF2_VARMIN;                       // 方差下限钳 / Variance floor
        END_IF
        _fInvA := DL_SF2_ONE / _fVarA;                     // A 逆方差（分母已钳底恒正） / Inverse variance of A
        _fInvB := DL_SF2_ONE / _fVarB;                     // B 逆方差 / Inverse variance of B
        _fW := _fInvA / (_fInvA + _fInvB);                 // 逆方差归一权重（分母两项恒正，无除零） / Normalized inverse-variance weight
        IF _fW < 0.0 THEN
            _fW := 0.0;                                    // 权重下钳 / Weight floor clamp
        END_IF
        IF _fW > DL_SF2_ONE THEN
            _fW := DL_SF2_ONE;                             // 权重上钳 / Weight ceiling clamp
        END_IF
        _fFused := _fW * fMeasA + (DL_SF2_ONE - _fW) * fMeasB;   // 加权融合 / Weighted fusion
        _fMean := _fFused;                                 // 更新递推参考点 / Update recursion reference
        bValid := TRUE;                                    // 双源融合有效 / Dual-source fusion valid
    ELSIF _bUseA THEN
        _fFused := fMeasA;                                 // 单源降级：全权重信 A（降级不拒算） / Degraded single source A
        _fMean := _fFused;                                 // 更新参考点 / Update reference
        _fW := DL_SF2_ONE;                                 // A 权重全一 / Full weight to A
        bValid := TRUE;                                    // 降级仍有效 / Degraded still valid
    ELSIF _bUseB THEN
        _fFused := fMeasB;                                 // 单源降级：全权重信 B / Degraded single source B
        _fMean := _fFused;                                 // 更新参考点 / Update reference
        _fW := 0.0;                                        // A 权重归零 / Zero weight to A
        bValid := TRUE;                                    // 降级仍有效 / Degraded still valid
    END_IF
    (* 双源同拍均不可用：无赋值分支 → _fFused/_fW 冻结上次值（规格②），bValid 保持 FALSE *)
END_IF

(* —— 段 3：出口单点映射（名实双出口同源，R191） —— *)
fFused   := _fFused;                                       // 融合值出口（失效期冻结） / Fused outlet, frozen on loss
fWeightA := _fW;                                           // 权重出口 / Weight outlet
bValid   := bValid AND (NOT _bErrLatch);                   // 有效标志（组态故障期强制无效） / Validity, forced invalid on fault
IF _bUseA AND _bUseB THEN
    bAgree := ABS(fMeasA - fMeasB) <= fDevMax;             // 双源一致性判据（浮点容差比较，禁 =） / Two-source agreement test
ELSE
    bAgree := TRUE;                                        // 单源降级无对可比：视为一致（诊断语义声明） / Single source: deemed consistent
END_IF
bError := _bErrLatch;                                      // 故障标志出口 / Error flag outlet

END_FUNCTION_BLOCK

(* ---- FB_DL_ShewhartRules.st ---- *)
(*==============================================================================
 * 组件名称 (Component)  : FB_DL_ShewhartRules
 * 所属子库 (Sublibrary) : DL_Algo
 * 当前版本 (Version)    : 1.0.0
 * 兼容性   (Platform)   : CODESYS 3.5+ / TwinCAT 3 / 汇川 InoProShop / 施耐德 Machine Expert
 *                         仅依赖 Standard.library（ABS），零厂商私有库
 * 功能描述 (Function)   : Shewhart 控制图判异位图（Western Electric/Nelson 8 条
 *                         判异准则，公开判据 clean-room 自实现，零文本移植）：
 *                           bit1 单点越 3σ ｜ bit2 连续 9 点同侧 CL
 *                           bit3 连续 6 点单调递升或递降 ｜ bit4 连续 14 点
 *                           交替升降 ｜ bit5 连续 3 点中 2 点越 2σ 同侧
 *                           bit6 连续 5 点中 4 点越 1σ 同侧 ｜ bit7 连续 15 点
 *                           在 1σ 带内 ｜ bit8 连续 8 点在 1σ 带外
 *                         z = (fSample − fCL) ÷ fSigma；连长计数 nRunLen（同侧
 *                         CL 连续点数，换侧归 1）；滚动历史窗 15 点（aZ 倒序
 *                         数组，[0] 最新），窗未填满只评低深度规则（边界防御，
 *                         规格指定）。复位清全部计数与历史。
 * 接口     (Interface)  : 输入 fSample 观测样本、fCL 中心线、fSigma 标准差
 *                         （域 > 0）、bReset 复位；输出 uRuleBits 判异位图
 *                         （bit1..bit8）、nRunLen 同侧连长 [点]、bAlarm 任一
 *                         判异命中、nFill 历史窗填充数（诊断透读）、eErrCode
 *                         错误码、bError 故障标志。
 * 边界     (Boundary)   : ① **属主边界（写死）：本件只做判异位图与连长计数，
 *                         不做控制限计算、不接管报警管理**；σ 估计归统计件。
 *                         ② 滚动窗边界防御：aZ 定长 0..14，入窗移位 FOR 自深
 *                         至浅（界宽常量 15，无越界）；规则 k 只在 nFill >= k
 *                         所需深度时评估（bit4 需 14 点、bit7 需 15 点，未填
 *                         满不评，防上电零历史假阳性）。
 *                         ③ 连长窗口滚动：换侧（z 符号变化）或 z=0 归 1；
 *                         同侧递增；bit2 = nRunLen >= 9。
 *                         ④ 非有限判据（R79 双判）：样本非有限 → 跳过入窗与
 *                         计数（窗口不污染），信息码 eSampleSkip，位图保持
 *                         上拍（锁存语义，非单拍抹除）。
 *                         ⑤ 组态闸：fSigma <= 0 或非有限 → 锁存故障 eCfgBad，
 *                         位图清零安全侧，解除沿 = bReset 上升沿（R45 配对）。
 *                         ⑥ 单调判据用严格不等号（相等点不打断单调链的口径
 *                         为「相等即中断」保守侧，头注释声明）。
 *                         ⑦ 零全局耦合（无 GVL / VAR_EXTERNAL / 物理地址）。
 * 分工声明 (Scope)      : 与 `FB_DL_CpkCalc`/`FB_DL_CpkIndex` 分工：过程能力
 *                         指数归那件、逐点判异归本件；与 `FB_DL_ParticleCounterStat`
 *                         分工：粒子计数统计归那件。
 * 来源标签 (Source Tag) : 自研线（Western Electric/Nelson 8 判异准则为公开 SPC
 *                         定义 clean-room 自实现，零文本移植）
 * 码表     (Codes)      : 本件不占用任何全局数字码位。出口为 WORD 位图 +
 *                         DINT 连长 + BOOL 组 + ENUM 错误码；数字码位待主控
 *                         收口阶段统一派号。
 * 红线自检 (Redline)    : R1 ✓ 零 GVL/VAR_EXTERNAL ｜ R2 ✓ 零 %I/%Q/%M ｜ R3 ✓ 纯 IEC 61131-3
 *                         R4 ✓ 窗界防御 + 除数前置闸 + 非有限跳过 + 组态锁存
 *                         ｜ R5 ✓ 声明逐行同行双语注释
 *                         R6 N/A（无 ENUM 状态机） ｜ R7 ✓ 一 R_TRIG 段 0 无条件刷新
 * 修订历史 (Revision)   : 2026-11-20  v1.0.0  R50 首版（批次 4 · 序号 16）
 * 验收向量 (Acceptance) : ① fCL=10, fSigma=1：单点 x=13.5 → z=3.5 > 3 →
 *                         uRuleBits.bit1=1，bAlarm=TRUE；② 连续 9 点
 *                         x=10.5（z=0.5 同侧）→ nRunLen=9，bit2=1；③ bit6：
 *                         最近 5 点 z=[1.2,1.1,1.4,1.0,1.3]（4 点 >=1）→
 *                         bit6=1；④ fSigma=0 → 锁存 eCfgBad；⑤ x=NaN →
 *                         eSampleSkip，窗不移位。
 *==============================================================================*)

(*-----------------------------------------------------------------------------
 * 枚举: E_DL_ShewErr（错误码；信息级不置 bError，故障级恒伴 bError=TRUE）
 *----------------------------------------------------------------------------*)
TYPE E_DL_ShewErr :
(
    eOk         := 0,   // 正常 / Normal
    eCfgBad     := 1,   // 故障级：fSigma 域非法（<=0 或非有限） / Fault: sigma illegal
    eSampleSkip := 2    // 信息级：样本非有限跳过，窗不移位 / Info: sample skipped, window held
);
END_TYPE

FUNCTION_BLOCK FB_DL_ShewhartRules
VAR_INPUT
    fSample : LREAL := 0.0;           // 观测样本 [工程单位] / Observed sample
    fCL     : LREAL := 0.0;           // 中心线 [工程单位] / Centre line
    fSigma  : LREAL := 1.0;           // 标准差，域 > 0 [工程单位] / Standard deviation
    bReset  : BOOL := FALSE;          // 复位，上升沿清位图/连长/历史窗全部计数 [-] / Reset clears all counters and window
END_VAR
VAR_OUTPUT
    uRuleBits : WORD;                 // 判异位图（bit1..bit8 对应 8 条准则） [-] / Rule bitmap, bits 1..8
    nRunLen   : DINT := 0;            // 同侧 CL 连长（换侧归 1） [点] / Same-side run length
    bAlarm    : BOOL;                 // 任一判异命中 [-] / Any rule hit
    nFill     : DINT := 0;            // 历史窗填充数（0..15，诊断透读） [点] / Window fill count
    eErrCode  : E_DL_ShewErr;         // 错误码出口 / Error code outlet
    bError    : BOOL;                 // 故障标志（组态锁存） [-] / Error flag, latched
END_VAR
VAR
    _aZ       : ARRAY[0..14] OF LREAL;   // z 值滚动历史窗（[0] 最新） [-] / Rolling z history window
    _uBits    : WORD;                 // 位图内部单源 / Bitmap internal source
    _nRun     : DINT := 0;            // 连长内部锁存 [点] / Run length latch
    _z        : LREAL;                // 当拍 z 分数 [-] / z score this scan
    _bSide    : BOOL;                 // 当拍样本在 CL 上侧（z > 0） [-] / Sample above CL
    _bSidePrev: BOOL := FALSE;        // 前拍样本侧别快照（换侧判据源） [-] / Previous sample side snapshot
    _bOk      : BOOL;                 // 当拍样本可入窗（有限 ∧ 无故障） [-] / Sample acceptable this scan
    _bNonFin  : BOOL;                 // 样本非有限当拍量 [-] / Sample non-finite
    _bCfgBad  : BOOL;                 // 组态非法当拍量 [-] / Illegal configuration
    _bErrLatch: BOOL;                 // 组态故障锁存位（解除沿 = bReset 上升沿） / Latched config fault
    _bAlt     : BOOL;                 // 交替升降判据中间量 [-] / Alternation test intermediate
    _nHi3     : DINT;                 // 最近 3 点越 2σ 上侧计数 [点] / Count beyond +2 sigma in last 3
    _nLo3     : DINT;                 // 最近 3 点越 2σ 下侧计数 [点] / Count beyond -2 sigma in last 3
    _nHi5     : DINT;                 // 最近 5 点越 1σ 上侧计数 [点] / Count beyond +1 sigma in last 5
    _nLo5     : DINT;                 // 最近 5 点越 1σ 下侧计数 [点] / Count beyond -1 sigma in last 5
    _bIn15    : BOOL;                 // 最近 15 点全在 1σ 带内 [-] / All 15 within 1 sigma
    _bOut8    : BOOL;                 // 最近 8 点全在 1σ 带外 [-] / All 8 beyond 1 sigma
    _bMonoUp  : BOOL;                 // 最近 6 点单调递升 [-] / Six points monotonic rising
    _bMonoDn  : BOOL;                 // 最近 6 点单调递降 [-] / Six points monotonic falling
    i         : DINT;                 // 窗循环索引 / Window loop index
    rtReset   : R_TRIG;               // 复位沿实例，段 0 无条件调用 / Reset edge instance
END_VAR
VAR CONSTANT
    DL_SHW_NWIN   : DINT  := 15;      // 历史窗定长 [点] / History window length
    DL_SHW_ZERO   : LREAL := 0.0;     // 判零基准 [-] / Zero base
    DL_SHW_SIG3   : LREAL := 3.0;     // bit1 判异倍率 [-] / Rule 1 sigma multiple
    DL_SHW_SIG2   : LREAL := 2.0;     // bit5 判异倍率 [-] / Rule 5 sigma multiple
    DL_SHW_SIG1   : LREAL := 1.0;     // bit6/7/8 判异倍率 [-] / Rule 6/7/8 sigma multiple
    DL_SHW_RUN9   : DINT  := 9;       // bit2 连长阈 [点] / Rule 2 run threshold
    DL_SHW_BIT1   : WORD  := 1;       // bit0 基准掩码（SHL 位移基准） [-] / Bit zero base mask
    DL_SHW_ZTOL   : LREAL := 1.0E-12; // 过零容差（|z| 低于此归换侧，禁浮点 = 判等） [-] / Zero-crossing tolerance
END_VAR

(* —— 段 0：组态闸 + 非有限判 + 沿刷新 —— *)
_bCfgBad := (fSigma <= DL_SHW_ZERO) OR (fSigma <> fSigma) OR ((fSigma - fSigma) <> DL_SHW_ZERO);   // σ 域闸（除数前置，R79 双判） / Sigma domain gate
_bNonFin := (fSample <> fSample) OR ((fSample - fSample) <> DL_SHW_ZERO);   // 样本非有限 / Sample non-finite
rtReset(CLK := bReset);               // 复位沿，每拍必调 / Reset edge, every scan

(* —— 段 1：复位沿（清位图/连长/填充数/历史窗全部计数，规格指定） —— *)
IF rtReset.Q THEN
    _bErrLatch := FALSE;              // 清组态锁存（R188 声明：解除沿 = bReset 上升沿） / Clear cfg latch
    _nRun := 0;                       // 清连长 / Clear run length
    nRunLen := 0;                     // 清连长出口 / Clear run outlet
    nFill := 0;                       // 清填充数 / Clear fill count
    _uBits := 0;                      // 清位图 / Clear bitmap
    FOR i := 0 TO (DL_SHW_NWIN - 1) DO
        _aZ[i] := DL_SHW_ZERO;        // 清历史窗 / Clear history window
    END_FOR
END_IF
IF _bCfgBad AND (NOT _bErrLatch) THEN
    _bErrLatch := TRUE;               // 锁存 / Latch
END_IF

(* —— 段 2：故障/正常分支分派（故障期位图安全侧清零、窗冻结） —— *)
IF _bErrLatch THEN
    _uBits := 0;                      // 故障安全侧位图清零（规格⑤） / Safe-side bitmap zero
ELSE
    _bOk := (NOT _bNonFin);           // 样本可入窗判据 / Sample acceptable
    IF _bOk THEN
        _uBits := 0;                  // 位图当拍重建（跳过拍保持上拍位图，规格④） / Rebuild bitmap on accepted samples
        _z := (fSample - fCL) / fSigma;   // z 分数（除数已闸，无除零） / z score
        _bSide := _z > DL_SHW_ZERO;   // 上侧判据（z=0 归换侧处理） / Above-CL test
        (* 滚动窗移位：自深至浅倒序拷贝，界宽常量 15 无越界 *)
        FOR i := (DL_SHW_NWIN - 1) TO 1 BY -1 DO
            _aZ[i] := _aZ[i - 1];     // 倒序拷贝 / Shift down
        END_FOR
        _aZ[0] := _z;                 // 最新样本入窗（唯一写入点） / Push newest
        IF nFill < DL_SHW_NWIN THEN
            nFill := nFill + 1;       // 填充数递增（上限 15） / Fill count up
        END_IF
        (* 连长计数：过零（容差）或换侧归 1，同侧递增 *)
        IF ABS(_z) < DL_SHW_ZTOL THEN
            _nRun := 1;               // 过零（|z| 低于容差）：连长归 1 / Zero crossing: reset to one
        ELSIF (nRunLen > 0) AND (_bSide <> _bSidePrev) THEN
            _nRun := 1;               // 换侧：连长归 1 / Side change: reset to one
        ELSE
            _nRun := nRunLen + 1;     // 首点（nRunLen=0）或同侧：递增 / First point or same side: increment
        END_IF
        nRunLen := _nRun;             // 连长落出口 / Run length outlet
        _bSidePrev := _bSide;         // 前拍侧别快照（下拍换侧判据源） / Side snapshot for next scan

        (* —— bit1：单点越 3σ —— *)
        IF ABS(_z) > DL_SHW_SIG3 THEN
            _uBits := _uBits OR SHL(DL_SHW_BIT1, 1);   // bit1 置位 / Set rule 1
        END_IF
        (* —— bit2：连续 9 点同侧 —— *)
        IF nRunLen >= DL_SHW_RUN9 THEN
            _uBits := _uBits OR SHL(DL_SHW_BIT1, 2);   // bit2 置位 / Set rule 2
        END_IF
        (* —— bit3：连续 6 点单调（相等即中断，保守侧，头注释⑥） —— *)
        IF nFill >= 6 THEN
            _bMonoUp := (_aZ[0] > _aZ[1]) AND (_aZ[1] > _aZ[2]) AND (_aZ[2] > _aZ[3])
                     AND (_aZ[3] > _aZ[4]) AND (_aZ[4] > _aZ[5]);   // 递升链 / Rising chain
            _bMonoDn := (_aZ[0] < _aZ[1]) AND (_aZ[1] < _aZ[2]) AND (_aZ[2] < _aZ[3])
                     AND (_aZ[3] < _aZ[4]) AND (_aZ[4] < _aZ[5]);   // 递降链 / Falling chain
            IF _bMonoUp OR _bMonoDn THEN
                _uBits := _uBits OR SHL(DL_SHW_BIT1, 3);   // bit3 置位 / Set rule 3
            END_IF
        END_IF
        (* —— bit4：连续 14 点交替升降（窗深 14） —— *)
        IF nFill >= 14 THEN
            _bAlt := TRUE;            // 交替判据起步 / Alternation preset
            FOR i := 1 TO 13 DO
                IF (( _aZ[i - 1] - _aZ[i]) * (_aZ[i] - _aZ[i + 1])) >= DL_SHW_ZERO THEN
                    _bAlt := FALSE;   // 相邻两差同号（含零差）：交替链断 / Same-sign diff: chain broken
                END_IF
            END_FOR
            IF _bAlt THEN
                _uBits := _uBits OR SHL(DL_SHW_BIT1, 4);   // bit4 置位 / Set rule 4
            END_IF
        END_IF
        (* —— bit5：最近 3 点中 2 点越 2σ 同侧 —— *)
        IF nFill >= 3 THEN
            _nHi3 := 0;               // 上侧计数清 / Hi count clear
            _nLo3 := 0;               // 下侧计数清 / Lo count clear
            FOR i := 0 TO 2 DO
                IF _aZ[i] >= DL_SHW_SIG2 THEN
                    _nHi3 := _nHi3 + 1;   // 越 +2σ 计数 / Count beyond +2 sigma
                ELSIF _aZ[i] <= (-DL_SHW_SIG2) THEN
                    _nLo3 := _nLo3 + 1;   // 越 -2σ 计数 / Count beyond -2 sigma
                END_IF
            END_FOR
            IF (_nHi3 >= 2) OR (_nLo3 >= 2) THEN
                _uBits := _uBits OR SHL(DL_SHW_BIT1, 5);   // bit5 置位 / Set rule 5
            END_IF
        END_IF
        (* —— bit6：最近 5 点中 4 点越 1σ 同侧 —— *)
        IF nFill >= 5 THEN
            _nHi5 := 0;               // 上侧计数清 / Hi count clear
            _nLo5 := 0;               // 下侧计数清 / Lo count clear
            FOR i := 0 TO 4 DO
                IF _aZ[i] >= DL_SHW_SIG1 THEN
                    _nHi5 := _nHi5 + 1;   // 越 +1σ 计数 / Count beyond +1 sigma
                ELSIF _aZ[i] <= (-DL_SHW_SIG1) THEN
                    _nLo5 := _nLo5 + 1;   // 越 -1σ 计数 / Count beyond -1 sigma
                END_IF
            END_FOR
            IF (_nHi5 >= 4) OR (_nLo5 >= 4) THEN
                _uBits := _uBits OR SHL(DL_SHW_BIT1, 6);   // bit6 置位 / Set rule 6
            END_IF
        END_IF
        (* —— bit7：连续 15 点在 1σ 带内（窗满才评） —— *)
        IF nFill >= DL_SHW_NWIN THEN
            _bIn15 := TRUE;           // 带内判据起步 / Within preset
            FOR i := 0 TO (DL_SHW_NWIN - 1) DO
                IF ABS(_aZ[i]) >= DL_SHW_SIG1 THEN
                    _bIn15 := FALSE;  // 任一点越带：判据断 / Any beyond band: broken
                END_IF
            END_FOR
            IF _bIn15 THEN
                _uBits := _uBits OR SHL(DL_SHW_BIT1, 7);   // bit7 置位 / Set rule 7
            END_IF
        END_IF
        (* —— bit8：连续 8 点在 1σ 带外 —— *)
        IF nFill >= 8 THEN
            _bOut8 := TRUE;           // 带外判据起步 / Beyond preset
            FOR i := 0 TO 7 DO
                IF ABS(_aZ[i]) < DL_SHW_SIG1 THEN
                    _bOut8 := FALSE;  // 任一点回带：判据断 / Any within band: broken
                END_IF
            END_FOR
            IF _bOut8 THEN
                _uBits := _uBits OR SHL(DL_SHW_BIT1, 8);   // bit8 置位 / Set rule 8
            END_IF
        END_IF
    END_IF
END_IF

(* —— 段 3：出口单点映射（名实双出口同源，R191） —— *)
uRuleBits := _uBits;                  // 位图出口 / Bitmap outlet
bAlarm := (_uBits <> 0);              // 任一判异命中 / Any rule hit
IF _bErrLatch THEN
    bError := TRUE;                   // 故障标志（R45 配对） / Error flag
    eErrCode := E_DL_ShewErr.eCfgBad; // 故障级码 / Fault code
ELSE
    bError := FALSE;                  // 无故障级条件 / No fault
    IF _bNonFin THEN
        eErrCode := E_DL_ShewErr.eSampleSkip;   // 信息级：样本跳过 / Info: skipped
    ELSE
        eErrCode := E_DL_ShewErr.eOk;           // 正常 / Normal
    END_IF
END_IF

END_FUNCTION_BLOCK

(* ---- FB_DL_SignalReconstruct.st ---- *)
(*==============================================================================
 * 组件名称 (Component)  : FB_DL_SignalReconstruct
 * 所属子库 (Sublibrary) : DL_Algo
 * 当前版本 (Version)    : 1.0.0
 * 兼容性 (Platform)     : CODESYS 3.5+ / TwinCAT 3 / 汇川 InoProShop / 施耐德 Machine Expert
 *                         仅依赖 Standard.library，零厂商私有库
 * 功能描述 (Function)   : 短丢包信号重构（状态估计族）。bSampleValid 电平指示
 *                         本拍采样有效；有效拍更新最近两次有效样本 (t1,v1)/(t2,v2)
 *                         并派生斜率 k = (v2-v1)/dt21；丢包期间按一阶外插
 *                         fOut = v2 + k·dtHold 输出，不确定度带按
 *                         fUncert = fUncBase + fUncRate·dtHold 随保持时长线性
 *                         增长（外插越久越不可信），bReconstructed 指示当前拍
 *                         为重构值。通信抖动、探头短时断流、HMI 采样缺口场景。
 * 来源标签 (Origin)     : 自研线（状态估计语义 clean-room，IEC 61131-3 标准语义的
 *                         道莅防御性实现，零代码行复制）
 * 边界语义 (Boundary)   : ① 丢 1 拍即可重构；连续丢包超过 tMaxHold → 停止外插，
 *                         bValid 强制 FALSE 并冻结末值（超窗重构比冻结更危险，
 *                         R133 语义：不把外推值伪装成测量）；
 *                         ② dt21 除零防御：两次有效样本间隔 <= eps → 斜率置 0
 *                         （零阶保持退化为常值外插），不产生 Inf；
 *                         ③ NaN 样本拒收：v1/v2 非有限 → 不入样本槽，bValid=FALSE；
 *                         ④ 组态闸：fUncBase < 0.0 或 fUncRate < 0.0 或
 *                         tMaxHold <= T#0S → 故障锁存。
 * 输出语义 (Fallback)   : 【R191】bValid = FALSE → fOut 冻结保持末次有效值
 *                         （不清零，避免下游把 0 当真值）；eFault 相 → 冻结 +
 *                         bError = TRUE。
 * 码位     (Codes)      : 按 R297 范式零 16# 码位硬编码；错误出口 BOOL+ENUM(eCause)，
 *                         码位待主控收口统一派号。
 * 红线自检 (Redline)    : 7 项红线已自检：R1 零全局 ✓｜R2 零物理地址 ✓｜R3 纯 IEC ✓
 *                         R4 除零防御（dt eps 闸）/NaN 拒收/组态闸 ✓
 *                         R5 双语同行注释 ✓｜R6 CASE 带 ELSE 兜底迁 eFault ✓
 *                         R7 无定时器实例（监视型），N/A ✓
 * 验收向量 (Acceptance) : V1 v1=10.0@t0、v2=12.0@t0+2s，丢包 1s 后
 *                         fOut=13.0（k=1/s 容差 1E-6）；
 *                         V2 丢包 3s（< tMaxHold=5s）→ fUncert = fUncBase + 3·fUncRate；
 *                         V3 连续丢包 6s（> 5s）→ bValid=FALSE 冻结末值。
 * 修订历史 (Revision)   : 2026-11-20  v1.0.0  R49 首版（批 2 · 序号 7）
 *==============================================================================*)
TYPE E_DL_SrcState :
(
    eIdle  := 0,                             (* 未取得首个有效样本（无基线可外插） / Idle, no baseline *)
    eRun   := 10,                            (* 样本流运行（有效拍更新 / 丢包拍外插） / Run: update or extrapolate *)
    eFault := 90                             (* 故障锁存相 / Fault latched phase *)
);
END_TYPE

TYPE E_DL_SrcCause :
(
    eNone       := 0,                        (* 无故障成因 / No cause *)
    eCfgIllegal := 1,                        (* 组态非法：不确定度参数越域 / Illegal config *)
    ePhaseBad   := 2                         (* 非法相位兜底 / Illegal phase fallback *)
);
END_TYPE

FUNCTION_BLOCK FB_DL_SignalReconstruct
VAR_INPUT
    fSample    : LREAL := 0.0;               (* 采样输入值 [工程单位] / Sample input value *)
    bSampleValid : BOOL := FALSE;            (* 本拍采样有效电平（通信链质量位直连）[-] / Sample-valid level this scan *)
    tScan      : TIME := T#100MS;            (* 扫描周期（保持时长积分步长），域 > T#0S [ms] / Scan cycle time step *)
    fUncBase   : LREAL := 0.1;               (* 不确定度基础项，域 >= 0.0 [工程单位] / Base uncertainty term *)
    fUncRate   : LREAL := 0.05;              (* 不确定度增长率，域 >= 0.0 [工程单位/s] / Uncertainty growth rate *)
    tMaxHold   : TIME := T#2S;               (* 最大允许外插保持时长，域 > T#0S [ms] / Max extrapolation hold time *)
    bEnable    : BOOL := TRUE;               (* 重构使能，FALSE 时冻结输出不外插 [-] / Enable *)
    bReset     : BOOL := FALSE;              (* 复位命令，上升沿清全部样本槽与锁存 [-] / Reset command *)
END_VAR
VAR_OUTPUT
    fOut          : LREAL;                   (* 重构/直通输出值（无效相冻结保持）[工程单位] / Output value *)
    fUncert       : LREAL;                   (* 当前不确定度带半宽 [工程单位] / Uncertainty band half-width *)
    bReconstructed: BOOL;                    (* 本拍为重构值（丢包外插拍）指示 [-] / Reconstructed-this-scan flag *)
    bValid        : BOOL;                    (* 输出可用性（超窗冻结时 FALSE）[-] / Output validity *)
    nHoldScans    : UDINT;                   (* 当前连续丢包拍数（诊断）[拍] / Consecutive hold scan count *)
    eState        : E_DL_SrcState;           (* 状态出口 / State outlet *)
    eCause        : E_DL_SrcCause;           (* 故障成因出口（R190 归因唯一） / Fault cause outlet *)
    bError        : BOOL;                    (* 故障锁存标志 [-] / Fault latch flag *)
END_VAR
VAR
    _eState  : E_DL_SrcState := E_DL_SrcState.eIdle;      (* 内部相位（CASE 唯一写入目标） / Internal phase *)
    _eCause  : E_DL_SrcCause := E_DL_SrcCause.eNone;      (* 故障成因锁存量 / Latched cause *)
    rtReset  : R_TRIG;                       (* 复位沿实例，段 0 无条件调用 / Reset edge instance *)
    _fV1     : LREAL;                        (* 基线样本 1 值（锁存槽）[工程单位] / Baseline sample 1 value *)
    _fV2     : LREAL;                        (* 基线样本 2 值（锁存槽）[工程单位] / Baseline sample 2 value *)
    _nT1     : UDINT;                        (* 样本 1 时间戳（扫描计数）[拍] / Sample 1 timestamp in scans *)
    _nT2     : UDINT;                        (* 样本 2 时间戳（扫描计数）[拍] / Sample 2 timestamp in scans *)
    _nScan   : UDINT;                        (* 全局扫描计数器（时间戳基）[拍] / Global scan counter *)
    _nHold   : UDINT;                        (* 连续丢包拍数锁存 [拍] / Consecutive hold count latch *)
    _fK      : LREAL;                        (* 外插斜率 = (v2-v1)/dt21 [工程单位/拍] / Extrapolation slope *)
    _fOutInt : LREAL;                        (* 内部输出保持槽（锁存量）[工程单位] / Internal output hold *)
    _bHave2  : BOOL;                         (* 已取得两个有效样本位（外插资格）[-] / Two-sample baseline acquired *)
    _bFault  : BOOL;                         (* 故障锁存位 / Latched fault bit *)
    _bCfgBad : BOOL;                         (* 组态非法当拍量 / Illegal config this scan *)
END_VAR
VAR CONSTANT
    DL_SRC_EPS : LREAL := 1.0E-9;            (* 样本间隔判零容差 [拍] / Sample-interval epsilon *)
END_VAR

(* —— 段 0：当拍判据派生 + 沿实例无条件刷新（R228A） —— *)
_bCfgBad := (fUncBase < 0.0) OR (fUncRate < 0.0) OR (tMaxHold <= T#0S) OR (tScan <= T#0S);   (* 组态闸覆盖每个域引脚（R151） / Config gate, every pin *)
rtReset(CLK := bReset);                                       (* 复位沿每拍必调 / Reset edge every scan *)
_nScan := _nScan + 1;                                         (* 扫描计数推进（UDINT 回绕：2^32 拍 @10ms ≈ 497 天，工程按期重启覆盖） / Scan counter advance *)

(* —— 段 1：单拍量预清零（R107） —— *)
bReconstructed := FALSE;                                      (* 重构指示预清，唯一分支置位 / Reconstructed flag preset *)
bValid := FALSE;                                              (* 有效性预清（派生出口，全路径赋值 R285） / Validity preset *)

(* —— 段 2：复位沿处理（作用域：清故障 + 清样本槽 + 清计数器 + 迁 eIdle，R283 逐项声明） —— *)
IF rtReset.Q THEN
    _bFault := FALSE;                                         (* 清故障锁存 / Clear fault *)
    _eCause := E_DL_SrcCause.eNone;                           (* 清成因 / Clear cause *)
    _fV1 := 0.0;                                              (* 清样本槽 1 / Clear slot 1 *)
    _fV2 := 0.0;                                              (* 清样本槽 2 / Clear slot 2 *)
    _nT1 := 0;                                                (* 清时间戳 1 / Clear timestamp 1 *)
    _nT2 := 0;                                                (* 清时间戳 2 / Clear timestamp 2 *)
    _nHold := 0;                                              (* 清丢包计数 / Clear hold count *)
    _nScan := 0;                                              (* 清时间戳基 / Clear timestamp base *)
    _fK := 0.0;                                               (* 清斜率 / Clear slope *)
    _fOutInt := 0.0;                                          (* 清输出保持槽 / Clear output hold *)
    _bHave2 := FALSE;                                         (* 清外插资格 / Clear baseline flag *)
    bValid := FALSE;                                          (* 输出有效性同步清 / Output validity clear *)
    _eState := E_DL_SrcState.eIdle;                           (* 迁待基线相 / Back to idle *)
END_IF

(* —— 段 3：组态闸故障锁存（R45 配对；锁存至复位沿，R189） —— *)
IF _bCfgBad AND NOT _bFault THEN
    _bFault := TRUE;                                          (* 锁存故障位 / Latch fault *)
    _eCause := E_DL_SrcCause.eCfgIllegal;                     (* 成因：组态非法 / Cause: illegal config *)
    _eState := E_DL_SrcState.eFault;                          (* 同步迁故障相 / Migrate to fault *)
END_IF

(* —— 段 4：CASE 主状态机（ELSE 兜底迁 eFault，红线 6） —— *)
CASE _eState OF
    E_DL_SrcState.eIdle:                                      (* 待基线相：只收样本不外插 / Idle: collect only *)
        IF bEnable AND NOT _bFault AND bSampleValid AND (fSample = fSample) AND ((fSample - fSample) = (fSample - fSample)) THEN
            _fV1 := fSample;                                  (* 首个有效样本入槽 1 / First sample into slot 1 *)
            _nT1 := _nScan;                                   (* 记时间戳 / Record timestamp *)
            _fOutInt := fSample;                              (* 直通输出 / Pass-through *)
            bValid := TRUE;                                   (* 单样本即可直通 / Valid with one sample *)
            _eState := E_DL_SrcState.eRun;                    (* 进入运行相 / Enter run *)
        END_IF
    E_DL_SrcState.eRun:                                       (* 运行相：有效拍更新 / 丢包拍外插 / Run *)
        IF NOT bEnable THEN                                   (* 失能：冻结输出（声明语义） / Disable: freeze *)
            _nHold := 0;                                      (* 清丢包计数 / Clear hold count *)
            _eState := E_DL_SrcState.eIdle;                   (* 回待基线（不重置样本槽，恢复使能即可续用基线） / Back to idle, slots kept *)
        ELSIF bSampleValid AND (fSample = fSample) AND ((fSample - fSample) = (fSample - fSample)) THEN
            (* 有效拍：旧 v2 滚动入 v1，新样本入 v2，斜率重派生 / Valid scan: roll slots, re-derive slope *)
            _fV1 := _fV2;                                     (* 槽 2 滚动入槽 1 / Roll slot 2 to slot 1 *)
            _nT1 := _nT2;                                     (* 时间戳同步滚动 / Roll timestamp *)
            _fV2 := fSample;                                  (* 新样本入槽 2 / New sample into slot 2 *)
            _nT2 := _nScan;                                   (* 新时间戳 / New timestamp *)
            IF (UDINT_TO_LREAL(_nT2 - _nT1)) > DL_SRC_EPS THEN
                _fK := (_fV2 - _fV1) / UDINT_TO_LREAL(_nT2 - _nT1);   (* 斜率派生：间隔已判非零，无除零 / Slope, divisor gated *)
            ELSE
                _fK := 0.0;                                   (* 同拍重复样本：斜率退化 0（零阶保持） / Degenerate slope zero *)
            END_IF
            _bHave2 := TRUE;                                  (* 外插资格确立 / Baseline acquired *)
            _fOutInt := fSample;                              (* 直通输出 / Pass-through *)
            fUncert := fUncBase;                              (* 有效拍不确定度 = 基础项 / Uncertainty = base *)
            _nHold := 0;                                      (* 清丢包计数 / Clear hold count *)
            bValid := TRUE;                                   (* 有效 / Valid *)
        ELSE
            (* 丢包拍：一阶外插 + 不确定度线性增长 / Dropped scan: extrapolate *)
            _nHold := _nHold + 1;                             (* 丢包计数递增 / Hold count advance *)
            _fOutInt := _fV2 + _fK * UDINT_TO_LREAL(_nHold);  (* 一阶外插（斜率按拍计） / First-order extrapolation *)
            fUncert := fUncBase + fUncRate * UDINT_TO_LREAL(_nHold) * TIME_TO_LREAL(tScan) / 1000.0;   (* 不确定度带：基础项 + 增长率·保持秒 / Uncertainty band growth *)
            IF _bHave2 THEN
                bValid := TRUE;                               (* 有基线：外插值有效 / Baseline: extrapolation valid *)
                bReconstructed := TRUE;                       (* 重构指示 / Reconstructed flag *)
            END_IF
            IF (tMaxHold > T#0S) AND (UDINT_TO_LREAL(_nHold) * TIME_TO_LREAL(tScan) / 1000.0 > TIME_TO_LREAL(tMaxHold) / 1000.0) THEN
                bValid := FALSE;                              (* 超窗：停止外插信任，冻结末值（R133 不伪装测量） / Beyond window: freeze, stop trusting extrapolation *)
                _fOutInt := _fV2;                             (* 冻结到末次有效样本 / Freeze to last valid sample *)
                fUncert := fUncBase + fUncRate * TIME_TO_LREAL(tMaxHold) / 1000.0;   (* 不确定度封顶在窗界 / Cap uncertainty at window bound *)
            END_IF
        END_IF
    E_DL_SrcState.eFault:                                     (* 故障相：冻结保持，仅复位沿出 / Fault *)
        ;                                                     (* 锁存回放（R28） / Replay from latch *)
    ELSE                                                      (* 非法相位兜底迁安全态 / Illegal phase fallback *)
        _eState := E_DL_SrcState.eFault;                      (* 迁故障相 / To fault *)
        _bFault := TRUE;                                      (* 同步锁存 / Latch *)
        _eCause := E_DL_SrcCause.ePhaseBad;                   (* 成因：非法相位 / Cause: illegal phase *)
END_CASE

(* —— 段 5：出口映射（bError/eState 同源，R191） —— *)
fOut := _fOutInt;                                             (* 输出单点映射 / Output mapping *)
nHoldScans := _nHold;                                         (* 丢包计数镜像 / Hold count mirror *)
bError := _bFault;                                            (* 故障标志镜像 / Fault flag mirror *)
eState := _eState;                                            (* 状态出口 / State outlet *)
eCause := _eCause;                                            (* 成因出口 / Cause outlet *)
END_FUNCTION_BLOCK

(* ---- FB_DL_SmithPredictor.st ---- *)
(*==============================================================================
 * 组件名称 (Component)  : FB_DL_SmithPredictor
 * 所属子库 (Sublibrary) : DL_Algo
 * 当前版本 (Version)    : 1.0.1
 * 兼容性   (Platform)   : CODESYS 3.5 / TwinCAT 3 / 汇川 InoProShop / Machine Expert
 *                         仅依赖 Standard.library（R_TRIG 经子块间接使用），零厂商方言
 * 功能描述 (Function)   : 大滞后对象专用史密斯预估器。内部按一阶 + 纯滞后模型
 *                         实时仿真"若无滞后过程会如何响应"，用补偿后误差驱动内
 *                         嵌 PID，等效消除纯滞后对环路稳定性的破坏；模型静态偏
 *                         差经小增益在线自适应校正。上电后队列填充期自动退化为
 *                         普通 PID（学习态），不阻塞控制。现场用途：长管道加热、
 *                         烘箱等大纯滞后温控回路。
 * 开源溯源 (Origin)     : 原创实现。史密斯预估器功能分类与参数域参考过程控制
 *                         经典文献（Smith dead-time compensator）的公开语义描
 *                         述，未复制任何厂商源码，clean-room 重写。
 * 本文件内含       : TYPE  E_DL_SmithState（配套枚举，归属 DL_Algo）
 *                    FB    FB_DL_SmithPredictor
 * 依赖     (Depends)    : FB_DL_PidController（DL_Algo 内部）
 * 红线自检 (Redline)    : R1 ✓ 零全局变量表与外部变量引用 ｜ R2 ✓ 零物理 IO 地址直写
 *                         R3 ✓ 纯 IEC 61131-3 ｜ R4 ✓ 防除零+钳位+数组边界防御
 *                         R5 ✓ 全变量中英双语同行注释 ｜ R6 ✓ 五态 ENUM+CASE+ELSE
 *                         R7 ✓ R_TRIG 实例主体最前部无条件刷新
 * 修订历史 (Revision)   :
 *   2026-11-15  v1.0.0  首版入库 · Round 04 · Level 1 DL_Algo
 *   2026-11-15  v1.0.1  阶段五终审精修：信息级码 0502（模型滞后截断）不再
 *                       置 bError，防下游报警误动作
 * 验收向量 (Acceptance) :
 *   V1 学习态：上电前 nLagSteps 拍内 fErrComp = fSetpoint - fPv（未补偿）
 *   V2 补偿态：队列填满后 fErrComp = fPv - (fModelDelayed + fModelBias)
 *   V3 模型收敛：fModelK=1, tModelT=T#1S, 恒定控制量 50 → fModelOut 趋近 50
 *   V4 自适应：对象静差存在 → fModelBias 朝消除偏差方向缓慢增长
 *   V5 增益非法：fModelK=0 → fModelOut 恒 0 且码 0002_0501，控制不中断
 *   V6 手动无扰：手动 30.0 切自动首拍输出保持 30.0 连续
 *============================================================================*)

(*-----------------------------------------------------------------------------
 * 枚举: E_DL_SmithState（归属 DL_Algo，与 FB_DL_SmithPredictor 同文件）
 * 含义: 史密斯预估器离散状态。数值步长留空位便于后续插态而不破坏已有工程。
 *----------------------------------------------------------------------------*)
TYPE E_DL_SmithState :
(
    eIdle         := 0,   // 使能关：模型与队列冻结，输出回下限 / Idle: model frozen, output at low limit
    eLearning     := 10,  // 学习态：队列填充中，PID 用原始误差 / Learning: queue filling, PID uses raw error
    eCompensating := 20,  // 补偿态：队列满，全补偿闭环 / Compensating: queue full, full compensation
    eManual       := 30,  // 手动态：输出手动值，模型继续仿真 / Manual: manual output, model still simulates
    eFault        := 99   // 故障兜底态：非法状态进入，输出安全值 / Fault fallback: illegal state, safe output
);
END_TYPE

(*==============================================================================
 * 功能块: FB_DL_SmithPredictor
 * 调用约定: 每个扫描周期无条件调用一次；bReset 上升沿重置模型与队列。
 * 无状态泄漏: 全部状态驻留于实例私有 VAR，零全局引用，可多实例并行。
 * 工程披露: 模型滞后队列为固定 20 槽环形缓冲，深度按 tModelLag/tSampleTime
 *           向下取整折算，超出上限截断并置码，不做动态扩容。
 *============================================================================*)
FUNCTION_BLOCK FB_DL_SmithPredictor
VAR_INPUT
    bEnable     : BOOL := FALSE;      // 总使能，FALSE 时输出回下限 / Master enable, FALSE drives output to low limit
    bManual     : BOOL := FALSE;      // 手动模式，TRUE 时输出手动值 / Manual mode, TRUE outputs manual value
    fManualValue: REAL := 0.0;        // 手动输出值 [%]，越限自动钳位 / Manual output value, auto-clamped
    fSetpoint   : REAL := 0.0;        // 设定值 [EU] / Setpoint in engineering units
    fPv         : REAL := 0.0;        // 过程值 [EU] / Process value in engineering units
    fKp         : REAL := 1.0;        // 内嵌 PID 比例增益 [1] / Embedded PID proportional gain
    tTi         : TIME := T#2S;       // 内嵌 PID 积分时间 [s] / Embedded PID integral time
    tTd         : TIME := T#0S;       // 内嵌 PID 微分时间 [s] / Embedded PID derivative time
    fModelK     : REAL := 1.0;        // 对象模型增益 [EU/EU] / Plant model gain
    tModelT     : TIME := T#5S;       // 模型惯性时间 [s] / Model time constant in seconds
    tModelLag   : TIME := T#1S;       // 模型纯滞后 [s] / Model dead time in seconds
    rOutMin     : REAL := 0.0;        // 输出下限 [%] / Output lower limit in percent
    rOutMax     : REAL := 100.0;      // 输出上限 [%] / Output upper limit in percent
    tSampleTime : TIME := T#100MS;    // 采样周期 [s] / Sample period in seconds
    bReset      : BOOL := FALSE;      // 复位信号，上升沿重置模型 / Reset, rising edge resets model
END_VAR
VAR_OUTPUT
    fCtrlOut    : REAL;               // 控制器输出 [%] / Controller output in percent
    fModelOut   : REAL;               // 模型无滞后输出 [EU]，诊断 / Model no-delay output, diagnostics
    fErrComp    : REAL;               // 补偿后偏差 [EU]，诊断 / Compensated error, diagnostics
    fModelBias  : REAL;               // 模型自适应偏差 [EU] / Model adaptive bias
    bError      : BOOL;               // 故障标志 / Fault flag
    uErrorId    : UDINT;              // 故障码，0 = 无故障 / Error code, 0 = no error
END_VAR
VAR
    fbPid       : FB_DL_PidController;  // 内嵌 PID 实例 / Embedded PID instance
    fModelState : REAL;               // 一阶模型状态 [EU] / First-order model state
    afLagBuf    : ARRAY[0..19] OF REAL;  // 模型滞后队列 [EU]，20 槽环形 / Model delay queue, 20-slot ring
    nLagSteps   : INT;                // 队列深度 = tModelLag/tSampleTime [拍] / Queue depth in cycles
    nWriteIdx   : INT;                // 环形队列写指针 [0..19] / Ring buffer write index
    nFillCnt    : INT;                // 队列填充计数 [拍] / Queue fill counter in cycles
    eState      : E_DL_SmithState;    // 主状态机当前状态 / Current state of the state machine
    bInit       : BOOL := FALSE;      // 首扫初始化标志 / First-scan init flag
    fbTrigReset : R_TRIG;             // 复位信号上升沿检测实例 / Reset rising edge detector instance
    fDt         : REAL;               // 生效采样周期 [s] / Effective sample period in seconds
    fLimLow     : REAL;               // 修复后的输出下限 [%] / Repaired output lower limit
    fLimHigh    : REAL;               // 修复后的输出上限 [%] / Repaired output upper limit
    fModelDelayed: REAL;              // 滞后队列读出的模型输出 [EU] / Delayed model output from queue
    fErrRaw     : REAL;               // 原始未补偿偏差 [EU] / Raw uncompensated error
    nReadIdx    : INT;                // 环形队列读指针 [0..19] / Ring buffer read index
    nDepthRaw   : INT;                // 折算的原始队列深度 [拍] / Raw computed queue depth in cycles
    bNonFinite  : BOOL;               // 本拍输入非有限值标志 / Non-finite input flag of this cycle
END_VAR
VAR CONSTANT
    DL_SMITH_LAG_MAX : INT  := 20;    // 模型滞后队列深度上限 [槽] / Model delay queue ceiling in slots
    DL_SMITH_KB      : REAL := 0.02;  // 模型偏差自适应增益 [1/s] / Model bias adaptive gain
END_VAR

(*------------------------------------------------------------------------------
 * 段 1｜无条件刷新区（红线 R7）：复位沿检测严禁进入任何 IF / CASE 分支
 *      Unconditional refresh zone (red line R7): edge detector outside IF / CASE
 *-----------------------------------------------------------------------------*)
fbTrigReset(CLK := bReset);

(*------------------------------------------------------------------------------
 * 段 2｜参数钳位与公共防御（不中断扫描）
 *      Parameter clamping and common defenses, never stops the scan
 *-----------------------------------------------------------------------------*)
bError   := FALSE;                    // 每拍重算故障标志 / Recompute fault flag every cycle
uErrorId := 16#0002_0000;             // 每拍重算故障码 / Recompute error code every cycle
bNonFinite := FALSE;                  // 非有限值标志每拍重算 / Non-finite flag recomputed every cycle

IF tSampleTime < T#10MS THEN
    fDt := 0.01;                      // 采样周期非法钳位为 0.01 s / Illegal sample period clamped to 0.01 s
    uErrorId := 16#0002_0002;         // 公共码：采样周期已钳位 / Common code: sample period clamped
ELSE
    fDt := TIME_TO_REAL(tSampleTime) / 1000.0;  // 采样周期换算为秒 [s] / Sample period in seconds
END_IF

IF rOutMin > rOutMax THEN
    fLimLow  := rOutMax;              // 上下限对调修复 / Swapped repair of limits
    fLimHigh := rOutMin;              // 上下限对调修复 / Swapped repair of limits
    uErrorId := 16#0002_0001;         // 公共码：参数越界已钳位 / Common code: parameter clamped
ELSE
    fLimLow  := rOutMin;              // 合法下限直通 / Valid low limit passed
    fLimHigh := rOutMax;              // 合法上限直通 / Valid high limit passed
END_IF

(* 模型滞后深度折算：向下取整，超上限截断置码 *)
(* Model lag depth derivation: floor division, truncated at ceiling with code *)
nDepthRaw := REAL_TO_INT(TRUNC(TIME_TO_REAL(tModelLag) / 1000.0 / fDt));  // 原始深度 [拍] / Raw depth in cycles
IF nDepthRaw > DL_SMITH_LAG_MAX THEN
    nLagSteps := DL_SMITH_LAG_MAX;    // 深度截断至上限 / Depth truncated to ceiling
    uErrorId := 16#0002_0502;         // 组件码：模型滞后超队列上限已截断 / Code: model lag truncated
ELSIF nDepthRaw < 0 THEN
    nLagSteps := 0;                   // 负深度防御为 0 / Negative depth defended to zero
ELSE
    nLagSteps := nDepthRaw;           // 合法深度直通 / Valid depth passed
END_IF

(* 模型增益非法防御：增益为 0 时模型输出恒 0，控制不中断 *)
(* Model gain defense: zero gain gives zero model output, control continues *)
IF fModelK = 0.0 THEN
    uErrorId := 16#0002_0501;         // 组件码：模型增益非法 / Code: model gain illegal
END_IF

(* 输入非有限值防御：设定或过程值非法即拒绝本拍更新 *)
(* Non-finite defense: reject this cycle if setpoint or process value invalid *)
IF (fSetpoint <> fSetpoint) OR (ABS(fSetpoint) > 1.0E30)
   OR (fPv <> fPv) OR (ABS(fPv) > 1.0E30)
   OR (fManualValue <> fManualValue) OR (ABS(fManualValue) > 1.0E30) THEN
    bNonFinite := TRUE;               // 置非有限值标志 / Set non-finite flag
END_IF

(*------------------------------------------------------------------------------
 * 段 3｜复位与首扫初始化：模型状态对齐过程值，队列预填，偏差清零
 *      Reset and first-scan init: model aligned to PV, queue prefilled
 *-----------------------------------------------------------------------------*)
IF fbTrigReset.Q OR (NOT bInit) THEN
    fModelState := fPv;               // 模型状态对齐过程值防上电冲击 / Model state aligned to PV
    fModelBias  := 0.0;               // 自适应偏差清零 / Adaptive bias cleared
    nWriteIdx   := 0;                 // 写指针归零 / Write index reset
    nFillCnt    := 0;                 // 填充计数归零 / Fill counter reset
    FOR nReadIdx := 0 TO DL_SMITH_LAG_MAX - 1 DO
        afLagBuf[nReadIdx] := fPv;    // 队列全槽预填过程值 / Prefill all queue slots with PV
    END_FOR
    bInit := TRUE;                    // 置首扫完成标志 / Set first-scan done flag
END_IF

IF NOT bEnable THEN
    eState  := eIdle;                 // 强制回空闲态 / Force idle state
    fCtrlOut:= fLimLow;               // 输出回下限 / Output to low limit
    RETURN;                           // 本拍结束（模型冻结） / End of cycle, model frozen
END_IF

IF bNonFinite THEN
    bError   := TRUE;                 // 置故障标志 / Set fault flag
    uErrorId := 16#0002_0004;         // 公共码：输入非有限值已拒绝 / Common code: non-finite rejected
    RETURN;                           // 保持上一拍输出与状态 / Hold previous output and state
END_IF

(*------------------------------------------------------------------------------
 * 段 4｜模型仿真：一阶惯性递推 + 增益折算 + 纯滞后队列 + 自适应偏差
 *      Model simulation: first-order recursion, gain scaling, queue, bias adaptation
 *-----------------------------------------------------------------------------*)
fModelState := fModelState + (fCtrlOut - fModelState) * fDt
               / MAX(TIME_TO_REAL(tModelT) / 1000.0, fDt);          // 一阶惯性递推 / First-order recursion
fModelOut := fModelState * fModelK;                                   // 增益折算输出 [EU] / Gain-scaled output

afLagBuf[nWriteIdx] := fModelOut;                                     // 当前模型输出入队 / Enqueue model output
nReadIdx := (nWriteIdx - nLagSteps + DL_SMITH_LAG_MAX) MOD DL_SMITH_LAG_MAX;  // 读指针 / Read index
nReadIdx := LIMIT(0, nReadIdx, DL_SMITH_LAG_MAX - 1);                 // 读指针防御钳位 / Defensive index clamp
fModelDelayed := afLagBuf[nReadIdx];                                  // 滞后读出 [EU] / Delayed readout
nWriteIdx := (nWriteIdx + 1) MOD DL_SMITH_LAG_MAX;                    // 写指针推进 / Advance write index

(* 队列填充计数：饱和于深度值，用于学习态判定 *)
(* Queue fill counter: saturated at depth, used for learning-state decision *)
IF nFillCnt < DL_SMITH_LAG_MAX THEN
    nFillCnt := nFillCnt + 1;         // 填充计数递增 / Increment fill counter
END_IF

(* 模型静态偏差在线自适应校正：小增益缓慢收敛 *)
(* Online adaptive bias correction: small gain slow convergence *)
fModelBias := fModelBias + DL_SMITH_KB * (fPv - fModelDelayed - fModelBias) * fDt;

(*------------------------------------------------------------------------------
 * 段 5｜内嵌 PID 引脚注入（本块不自写 PID 律）
 *      Embedded PID pin injection, no PID law rewritten here
 *-----------------------------------------------------------------------------*)
fbPid.bEnable      := TRUE;           // PID 使能 / PID enabled
fbPid.fSetpoint    := fErrComp;       // 设定 = 补偿后误差（实际引脚恒 0）/ Setpoint equals compensated error
fbPid.fActual      := 0.0;            // 实际恒 0，使偏差 = 补偿误差 / Actual zero so error equals compensated error
fbPid.fKp          := fKp;            // 增益透传 / Gain passthrough
fbPid.tTi          := tTi;            // 积分时间透传 / Integral time passthrough
fbPid.tTd          := tTd;            // 微分时间透传 / Derivative time passthrough
fbPid.fDeadband    := 0.0;            // 死区默认关闭 / Deadband off by default
fbPid.bIncremental := FALSE;          // 默认位置式 / Positional by default
fbPid.rOutMin      := rOutMin;        // 输出下限透传 / Low limit passthrough
fbPid.rOutMax      := rOutMax;        // 输出上限透传 / High limit passthrough
fbPid.tSampleTime  := tSampleTime;   // 采样周期透传 / Sample period passthrough
fbPid.bTrack       := FALSE;          // PID 自身不跟踪 / PID tracking off
fbPid.fTrackValue  := 0.0;            // 跟踪值占位 / Track value placeholder
fbPid.bReset       := bReset;         // 复位透传 / Reset passthrough

(*------------------------------------------------------------------------------
 * 段 6｜主状态机（红线 R6）：ENUM + CASE + ELSE 兜底
 *      Main state machine: ENUM + CASE with mandatory ELSE fallback
 *-----------------------------------------------------------------------------*)
CASE eState OF

    eIdle:
        (* 空闲态已在早退段处理；本分支仅做迁移防御 *)
        (* Idle handled in early exit; this branch only guards transfers *)
        IF bEnable THEN
            IF bManual THEN
                eState := eManual;    // 请求手动 / Request manual mode
            ELSIF nFillCnt < nLagSteps THEN
                eState := eLearning;  // 队列未满进学习态 / Queue not full, learning state
            ELSE
                eState := eCompensating;  // 队列满进补偿态 / Queue full, compensating
            END_IF
        END_IF

    eLearning:
        (* 学习态：队列填充中，PID 用原始误差闭环，不阻塞控制 *)
        (* Learning: queue filling, PID closed loop on raw error, control not blocked *)
        fErrRaw  := fSetpoint - fPv;  // 原始偏差 [EU] / Raw error
        fErrComp := fErrRaw;          // 补偿误差 = 原始误差 / Compensated equals raw
        fbPid.fSetpoint := fErrComp;  // 设定 = 补偿后误差 / Setpoint equals compensated error
        fbPid.bManual := FALSE;       // PID 自动 / PID auto
        fbPid();                      // PID 运算 / PID computation
        fCtrlOut := fbPid.fOut;       // 输出透传 / Output passthrough
        IF bManual THEN
            eState := eManual;        // 切手动 / Switch to manual
        ELSIF nFillCnt >= nLagSteps THEN
            eState := eCompensating;  // 队列满切补偿 / Queue full, compensating
        END_IF

    eCompensating:
        (* 补偿态：用模型滞后输出与自适应偏差重构等效无滞后误差 *)
        (* Compensating: reconstruct delay-free error from delayed model and bias *)
        fErrComp := fPv - (fModelDelayed + fModelBias);   // 补偿后偏差 [EU] / Compensated error
        fbPid.fSetpoint := fErrComp;  // 设定 = 补偿后误差 / Setpoint equals compensated error
        fbPid.bManual := FALSE;       // PID 自动 / PID auto
        fbPid();                      // PID 运算 / PID computation
        fCtrlOut := fbPid.fOut;       // 输出透传 / Output passthrough
        IF bManual THEN
            eState := eManual;        // 切手动 / Switch to manual
        END_IF

    eManual:
        (* 手动态：输出手动值（钳位），模型与队列继续仿真保证回自动连续 *)
        (* Manual: clamped manual output, model keeps simulating for bumpless return *)
        fErrRaw  := fSetpoint - fPv;  // 原始偏差诊断 / Raw error diagnostics
        fErrComp := fErrRaw;          // 补偿误差诊断 / Compensated error diagnostics
        fbPid.bManual     := TRUE;    // PID 手动 / PID manual
        fbPid.fManualValue:= fManualValue;  // 手动值注入 / Inject manual value
        fbPid();                      // PID 手动运算 / PID manual computation
        fbPid.bManual     := FALSE;   // 恢复自动配置位 / Restore auto config bit
        fCtrlOut := fbPid.fOut;       // 输出透传 / Output passthrough
        IF NOT bEnable THEN
            eState := eIdle;          // 切空闲 / Switch to idle
        ELSIF NOT bManual THEN
            IF nFillCnt >= nLagSteps THEN
                eState := eCompensating;  // 回补偿态 / Back to compensating
            ELSE
                eState := eLearning;  // 回学习态 / Back to learning
            END_IF
        END_IF

    eFault:
        (* 故障兜底态：输出安全下限，模型继续仿真 *)
        (* Fault fallback: safe low-limit output, model keeps simulating *)
        fCtrlOut := fLimLow;          // 安全输出 / Safe output

    ELSE
        (* 非法状态拦截：任何未定义状态一律进故障兜底，不做隐式恢复 *)
        (* Illegal state interception: any undefined state goes to fault fallback *)
        eState   := eFault;           // 进故障态 / Enter fault state
        bError   := TRUE;             // 置故障标志 / Set fault flag
        uErrorId := 16#0002_0005;     // 非法状态兜底码 / Illegal state fallback code
        fCtrlOut := fLimLow;          // 安全输出 / Safe output
END_CASE;

(* 信息级码（0502 模型滞后截断）不置故障标志，防下游报警误动作 *)
(* Info-level code (model lag truncation 0502) never raises the fault flag *)
bError := (uErrorId <> 16#0002_0000) AND (uErrorId <> 16#0002_0502);  // 非信息级码才置故障 / Fault flag only on non-info codes
END_FUNCTION_BLOCK
